REGION Network 2: Converstion all data to string
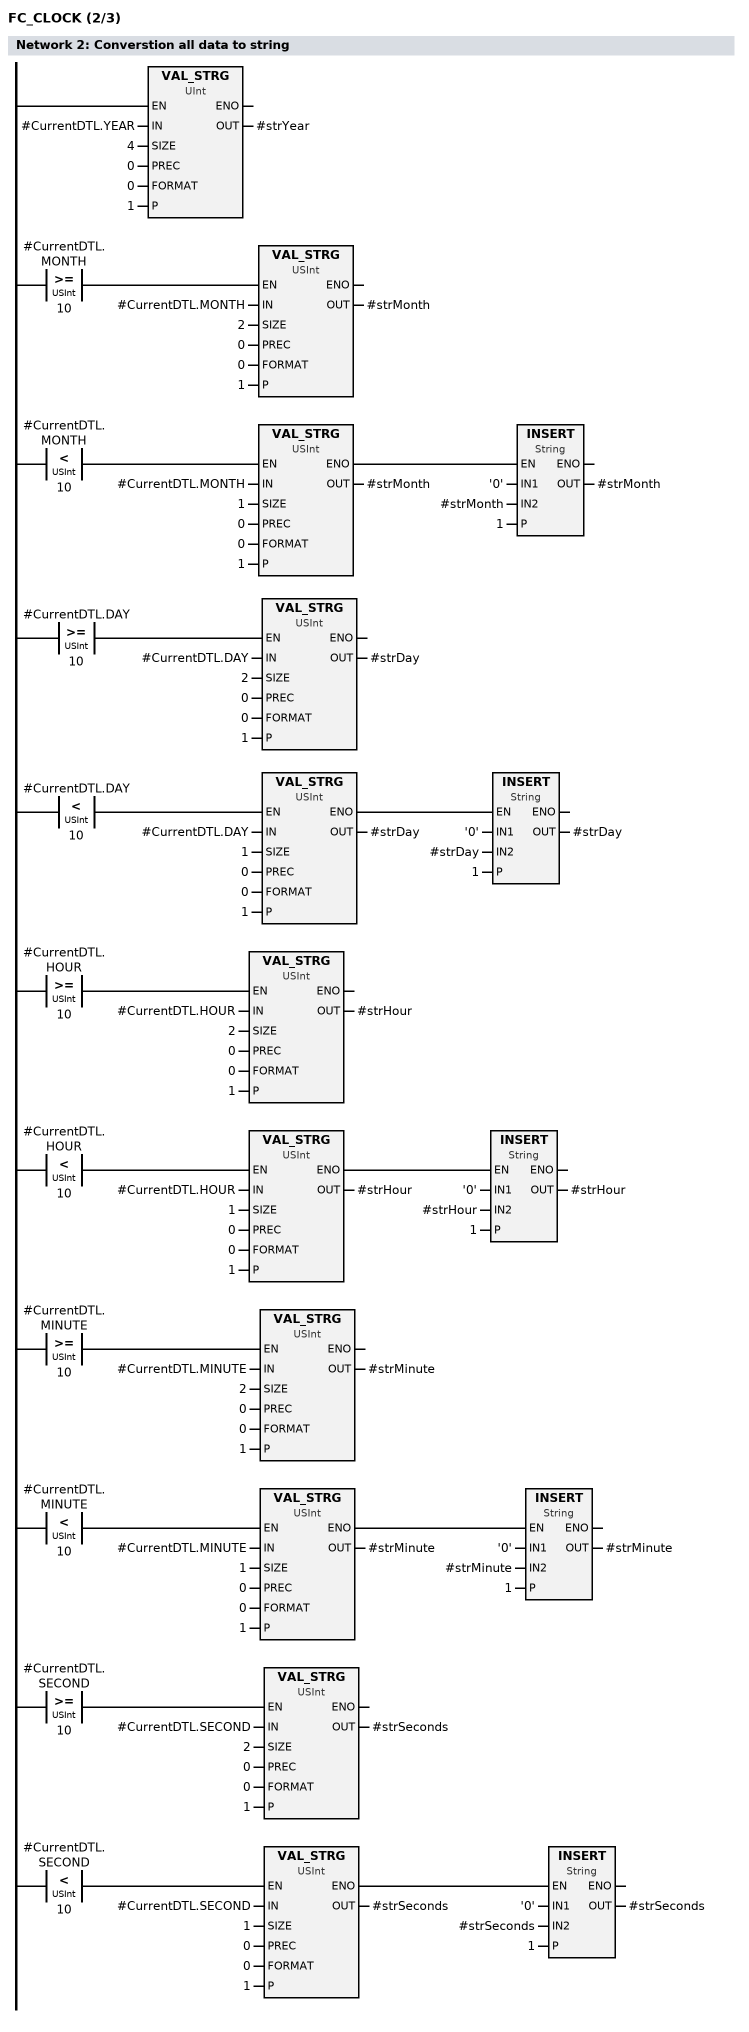
   RUNG wire#powerrail
      { S7_Templates := "[value_type := UInt, str_type := String]" } VAL_STRG(IN := #CurrentDTL.YEAR, SIZE := 4, PREC := 0, FORMAT := 0, P := 1, OUT => #strYear)
   END_RUNG
   RUNG wire#powerrail
      { S7_Templates := "SrcType := USInt" } GE_Contact(in1 := #CurrentDTL.MONTH, in2 := 10)
      { S7_Templates := "[value_type := USInt, str_type := String]" } VAL_STRG(IN := #CurrentDTL.MONTH, SIZE := 2, PREC := 0, FORMAT := 0, P := 1, OUT => #strMonth)
   END_RUNG
   RUNG wire#powerrail
      { S7_Templates := "SrcType := USInt" } LT_Contact(in1 := #CurrentDTL.MONTH, in2 := 10)
      { S7_Templates := "[value_type := USInt, str_type := String]" } VAL_STRG(IN := #CurrentDTL.MONTH, SIZE := 1, PREC := 0, FORMAT := 0, P := 1, OUT => #strMonth)
      { S7_Templates := "str_type := String" } INSERT(IN1 := '0', IN2 := #strMonth, P := 1, OUT => #strMonth)
   END_RUNG
   RUNG wire#powerrail
      { S7_Templates := "SrcType := USInt" } GE_Contact(in1 := #CurrentDTL.DAY, in2 := 10)
      { S7_Templates := "[value_type := USInt, str_type := String]" } VAL_STRG(IN := #CurrentDTL.DAY, SIZE := 2, PREC := 0, FORMAT := 0, P := 1, OUT => #strDay)
   END_RUNG
   RUNG wire#powerrail
      { S7_Templates := "SrcType := USInt" } LT_Contact(in1 := #CurrentDTL.DAY, in2 := 10)
      { S7_Templates := "[value_type := USInt, str_type := String]" } VAL_STRG(IN := #CurrentDTL.DAY, SIZE := 1, PREC := 0, FORMAT := 0, P := 1, OUT => #strDay)
      { S7_Templates := "str_type := String" } INSERT(IN1 := '0', IN2 := #strDay, P := 1, OUT => #strDay)
   END_RUNG
   RUNG wire#powerrail
      { S7_Templates := "SrcType := USInt" } GE_Contact(in1 := #CurrentDTL.HOUR, in2 := 10)
      { S7_Templates := "[value_type := USInt, str_type := String]" } VAL_STRG(IN := #CurrentDTL.HOUR, SIZE := 2, PREC := 0, FORMAT := 0, P := 1, OUT => #strHour)
   END_RUNG
   RUNG wire#powerrail
      { S7_Templates := "SrcType := USInt" } LT_Contact(in1 := #CurrentDTL.HOUR, in2 := 10)
      { S7_Templates := "[value_type := USInt, str_type := String]" } VAL_STRG(IN := #CurrentDTL.HOUR, SIZE := 1, PREC := 0, FORMAT := 0, P := 1, OUT => #strHour)
      { S7_Templates := "str_type := String" } INSERT(IN1 := '0', IN2 := #strHour, P := 1, OUT => #strHour)
   END_RUNG
   RUNG wire#powerrail
      { S7_Templates := "SrcType := USInt" } GE_Contact(in1 := #CurrentDTL.MINUTE, in2 := 10)
      { S7_Templates := "[value_type := USInt, str_type := String]" } VAL_STRG(IN := #CurrentDTL.MINUTE, SIZE := 2, PREC := 0, FORMAT := 0, P := 1, OUT => #strMinute)
   END_RUNG
   RUNG wire#powerrail
      { S7_Templates := "SrcType := USInt" } LT_Contact(in1 := #CurrentDTL.MINUTE, in2 := 10)
      { S7_Templates := "[value_type := USInt, str_type := String]" } VAL_STRG(IN := #CurrentDTL.MINUTE, SIZE := 1, PREC := 0, FORMAT := 0, P := 1, OUT => #strMinute)
      { S7_Templates := "str_type := String" } INSERT(IN1 := '0', IN2 := #strMinute, P := 1, OUT => #strMinute)
   END_RUNG
   RUNG wire#powerrail
      { S7_Templates := "SrcType := USInt" } GE_Contact(in1 := #CurrentDTL.SECOND, in2 := 10)
      { S7_Templates := "[value_type := USInt, str_type := String]" } VAL_STRG(IN := #CurrentDTL.SECOND, SIZE := 2, PREC := 0, FORMAT := 0, P := 1, OUT => #strSeconds)
   END_RUNG
   RUNG wire#powerrail
      { S7_Templates := "SrcType := USInt" } LT_Contact(in1 := #CurrentDTL.SECOND, in2 := 10)
      { S7_Templates := "[value_type := USInt, str_type := String]" } VAL_STRG(IN := #CurrentDTL.SECOND, SIZE := 1, PREC := 0, FORMAT := 0, P := 1, OUT => #strSeconds)
      { S7_Templates := "str_type := String" } INSERT(IN1 := '0', IN2 := #strSeconds, P := 1, OUT => #strSeconds)
   END_RUNG
   // the same network as SCL:
   VAL_STRG(IN := #CurrentDTL.YEAR, SIZE := 4, PREC := 0, FORMAT := 0, P := 1, OUT => #strYear);
   IF #CurrentDTL.MONTH >= 10 THEN
       VAL_STRG(IN := #CurrentDTL.MONTH, SIZE := 2, PREC := 0, FORMAT := 0, P := 1, OUT => #strMonth);
   END_IF;
   VAL_STRG(EN := #CurrentDTL.MONTH < 10,
            IN := #CurrentDTL.MONTH,
            SIZE := 1,
            PREC := 0,
            FORMAT := 0,
            P := 1,
            OUT => #strMonth,
            ENO => #_w1);
   IF #_w1 THEN INSERT(IN1 := '0', IN2 := #strMonth, P := 1, OUT => #strMonth); END_IF;
   IF #CurrentDTL.DAY >= 10 THEN
       VAL_STRG(IN := #CurrentDTL.DAY, SIZE := 2, PREC := 0, FORMAT := 0, P := 1, OUT => #strDay);
   END_IF;
   VAL_STRG(EN := #CurrentDTL.DAY < 10,
            IN := #CurrentDTL.DAY,
            SIZE := 1,
            PREC := 0,
            FORMAT := 0,
            P := 1,
            OUT => #strDay,
            ENO => #_w2);
   IF #_w2 THEN INSERT(IN1 := '0', IN2 := #strDay, P := 1, OUT => #strDay); END_IF;
   IF #CurrentDTL.HOUR >= 10 THEN
       VAL_STRG(IN := #CurrentDTL.HOUR, SIZE := 2, PREC := 0, FORMAT := 0, P := 1, OUT => #strHour);
   END_IF;
   VAL_STRG(EN := #CurrentDTL.HOUR < 10,
            IN := #CurrentDTL.HOUR,
            SIZE := 1,
            PREC := 0,
            FORMAT := 0,
            P := 1,
            OUT => #strHour,
            ENO => #_w3);
   IF #_w3 THEN INSERT(IN1 := '0', IN2 := #strHour, P := 1, OUT => #strHour); END_IF;
   IF #CurrentDTL.MINUTE >= 10 THEN
       VAL_STRG(IN := #CurrentDTL.MINUTE, SIZE := 2, PREC := 0, FORMAT := 0, P := 1, OUT => #strMinute);
   END_IF;
   VAL_STRG(EN := #CurrentDTL.MINUTE < 10,
            IN := #CurrentDTL.MINUTE,
            SIZE := 1,
            PREC := 0,
            FORMAT := 0,
            P := 1,
            OUT => #strMinute,
            ENO => #_w4);
   IF #_w4 THEN INSERT(IN1 := '0', IN2 := #strMinute, P := 1, OUT => #strMinute); END_IF;
   IF #CurrentDTL.SECOND >= 10 THEN
       VAL_STRG(IN := #CurrentDTL.SECOND, SIZE := 2, PREC := 0, FORMAT := 0, P := 1, OUT => #strSeconds);
   END_IF;
   VAL_STRG(EN := #CurrentDTL.SECOND < 10,
            IN := #CurrentDTL.SECOND,
            SIZE := 1,
            PREC := 0,
            FORMAT := 0,
            P := 1,
            OUT => #strSeconds,
            ENO => #_w5);
   IF #_w5 THEN INSERT(IN1 := '0', IN2 := #strSeconds, P := 1, OUT => #strSeconds); END_IF;
END_REGION

REGION Network 3: Current Time String
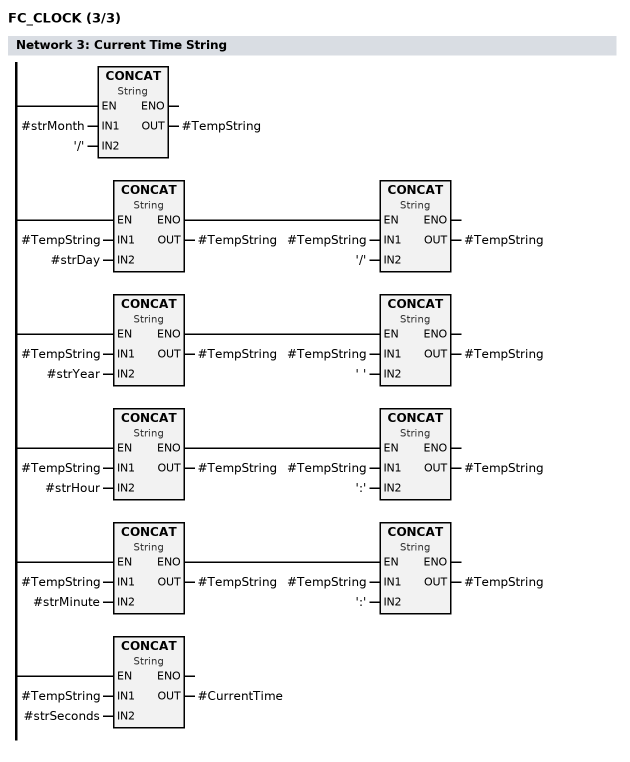
   RUNG wire#powerrail
      { S7_Templates := "[card := 2, str_type := String]" } CONCAT(IN1 := #strMonth, IN2 := '/', OUT => #TempString)
   END_RUNG
   RUNG wire#powerrail
      { S7_Templates := "[card := 2, str_type := String]" } CONCAT(IN1 := #TempString, IN2 := #strDay, OUT => #TempString)
      { S7_Templates := "[card := 2, str_type := String]" } CONCAT(IN1 := #TempString, IN2 := '/', OUT => #TempString)
   END_RUNG
   RUNG wire#powerrail
      { S7_Templates := "[card := 2, str_type := String]" } CONCAT(IN1 := #TempString, IN2 := #strYear, OUT => #TempString)
      { S7_Templates := "[card := 2, str_type := String]" } CONCAT(IN1 := #TempString, IN2 := ' ', OUT => #TempString)
   END_RUNG
   RUNG wire#powerrail
      { S7_Templates := "[card := 2, str_type := String]" } CONCAT(IN1 := #TempString, IN2 := #strHour, OUT => #TempString)
      { S7_Templates := "[card := 2, str_type := String]" } CONCAT(IN1 := #TempString, IN2 := ':', OUT => #TempString)
   END_RUNG
   RUNG wire#powerrail
      { S7_Templates := "[card := 2, str_type := String]" } CONCAT(IN1 := #TempString, IN2 := #strMinute, OUT => #TempString)
      { S7_Templates := "[card := 2, str_type := String]" } CONCAT(IN1 := #TempString, IN2 := ':', OUT => #TempString)
   END_RUNG
   RUNG wire#powerrail
      { S7_Templates := "[card := 2, str_type := String]" } CONCAT(IN1 := #TempString, IN2 := #strSeconds, OUT => #CurrentTime)
   END_RUNG
   // the same network as SCL:
   CONCAT(IN1 := #strMonth, IN2 := '/', OUT => #TempString);
   CONCAT(IN1 := #TempString, IN2 := #strDay, OUT => #TempString, ENO => #_w1);
   IF #_w1 THEN CONCAT(IN1 := #TempString, IN2 := '/', OUT => #TempString); END_IF;
   CONCAT(IN1 := #TempString, IN2 := #strYear, OUT => #TempString, ENO => #_w2);
   IF #_w2 THEN CONCAT(IN1 := #TempString, IN2 := ' ', OUT => #TempString); END_IF;
   CONCAT(IN1 := #TempString, IN2 := #strHour, OUT => #TempString, ENO => #_w3);
   IF #_w3 THEN CONCAT(IN1 := #TempString, IN2 := ':', OUT => #TempString); END_IF;
   CONCAT(IN1 := #TempString, IN2 := #strMinute, OUT => #TempString, ENO => #_w4);
   IF #_w4 THEN CONCAT(IN1 := #TempString, IN2 := ':', OUT => #TempString); END_IF;
   CONCAT(IN1 := #TempString, IN2 := #strSeconds, OUT => #CurrentTime);
END_REGION
END_FUNCTION

FUNCTION_BLOCK "FB_HeartBeat"   // FB25, SCL
{ S7_Optimized_Access := 'TRUE' }
VERSION : 0.1
// stored: AutoNumber true, IsIECCheckEnabled false, IsRetainMemResEnabled false, MemoryReserve 100, SetENOAutomatically false, UDAEnableTagReadback false
   VAR_INPUT
      PC_HeartBeat : Word;
   END_VAR
   VAR_OUTPUT
      PLC_HeartBeat : Word;
      PC_Disconnected : Bool;
   END_VAR
   VAR
      TimeOut : TON_TIME;
      "Timer" { S7_SetPoint := 'True'} : TON_TIME;
      PC_Heartbeat_old : Word;
      StartTimerBit : Bool := FALSE;
   END_VAR
BEGIN
   #Timer(IN := #StartTimerBit, //
          PT := t#250ms);
   IF NOT #StartTimerBit THEN
       #StartTimerBit := TRUE;
   END_IF;
   #Timer(IN := #StartTimerBit, //
          PT := t#250ms);
   IF #Timer.Q THEN
       #StartTimerBit := FALSE;
       RESET_TIMER(#Timer);
       #PLC_HeartBeat += 1;
   END_IF;
   //Time Out Timer
   #TimeOut(IN := #PC_HeartBeat = #PC_Heartbeat_old,
            PT := t#10s);
   #PC_Heartbeat_old := #PC_HeartBeat;
   #PC_Disconnected := #TimeOut.Q; // if time out set PC_Disconnected
END_FUNCTION_BLOCK

FUNCTION "OUTPUTS" : Void   // FC5, SCL
{ S7_Optimized_Access := 'TRUE' }
VERSION : 0.1
// stored: AutoNumber true, IsIECCheckEnabled false, SetENOAutomatically false, UDAEnableTagReadback false
BEGIN
   REGION MAIN PANEL
       "MAIN PANEL STACK LIGHT RED" := "Stack_Lights_DB_0".Red XOR "Force"."MAIN PANEL STACK LIGHT RED";
       "MAIN PANEL STACK LIGHT AMBER" := "Stack_Lights_DB_0".Yellow XOR "Force"."MAIN PANEL STACK LIGHT AMBER";
       "MAIN PANEL STACK LIGHT GREEN" := "Stack_Lights_DB_0".Green XOR "Force"."MAIN PANEL STACK LIGHT GREEN";
   END_REGION

   REGION REMOTE PANEL 1
       "C1101_SFTY STOPPER ROTATE" := "Sf_C1101_FB_DB".T_Run.Q XOR "Force".Remote_Panel[1]."CX101_SFTY STOPPER ROTATE";
       "C1102_SFTY STOPPER ROTATE" := "Sf_C1102_FB_DB".T_Run.Q XOR "Force".Remote_Panel[1]."CX102_SFTY STOPPER ROTATE";
       "C1103_SFTY STOPPER ROTATE" := "Sf_C1103_FB_DB".T_Run.Q XOR "Force".Remote_Panel[1]."CX103_SFTY STOPPER ROTATE";
       "C1104_SFTY STOPPER ROTATE" := "Sf_C1104_FB_DB".T_Run.Q XOR "Force".Remote_Panel[1]."CX104_SFTY STOPPER ROTATE";
       "C1105_SFTY STOPPER ROTATE" := "Sf_C1105_FB_DB".T_Run.Q XOR "Force".Remote_Panel[1]."CX105_SFTY STOPPER ROTATE";
       "C1106_SFTY STOPPER ROTATE" := "Sf_C1106_FB_DB".T_Run.Q XOR "Force".Remote_Panel[1]."CX106_SFTY STOPPER ROTATE";
       "C1107_SFTY STOPPER ROTATE" := "Sf_C1107_FB_DB".T_Run.Q XOR "Force".Remote_Panel[1]."CX107_SFTY STOPPER ROTATE";
       "C1108_SFTY STOPPER ROTATE" := "Sf_C1108_FB_DB".T_Run.Q XOR "Force".Remote_Panel[1]."CX108_SFTY STOPPER ROTATE";
       "C1201_SFTY STOPPER ROTATE" := "Sf_C1201_FB_DB".T_Run.Q XOR "Force".Remote_Panel[1]."CX201_SFTY STOPPER ROTATE";
       "C1202_SFTY STOPPER ROTATE" := "Sf_C1202_FB_DB".T_Run.Q XOR "Force".Remote_Panel[1]."CX202_SFTY STOPPER ROTATE";
       "C1203_SFTY STOPPER ROTATE" := "Sf_C1203_FB_DB".T_Run.Q XOR "Force".Remote_Panel[1]."CX203_SFTY STOPPER ROTATE";
       "C1204_SFTY STOPPER ROTATE" := "Sf_C1204_FB_DB".T_Run.Q XOR "Force".Remote_Panel[1]."CX204_SFTY STOPPER ROTATE";
       "C1205_SFTY STOPPER ROTATE" := "Sf_C1205_FB_DB".T_Run.Q XOR "Force".Remote_Panel[1]."CX205_SFTY STOPPER ROTATE";
       "C1206_SFTY STOPPER ROTATE" := "Sf_C1206_FB_DB".T_Run.Q XOR "Force".Remote_Panel[1]."CX206_SFTY STOPPER ROTATE";
       "C1207_SFTY STOPPER ROTATE" := "Sf_C1207_FB_DB".T_Run.Q XOR "Force".Remote_Panel[1]."CX207_SFTY STOPPER ROTATE";
       "C1208_SFTY STOPPER ROTATE" := "Sf_C1208_FB_DB".T_Run.Q XOR "Force".Remote_Panel[1]."CX208_SFTY STOPPER ROTATE";
       "VTD1 DOCKING PINS 1 EXTEND" := "Control_DB".VTD_Sys[1].Outputs.LP1_Extend XOR "Force".Remote_Panel[1]."VTDx DOCKING PINS 1 EXTEND";
       "VTD1 DOCKING PINS 1 RETRACT" := "Control_DB".VTD_Sys[1].Outputs.LP1_Retract XOR "Force".Remote_Panel[1]."VTDx DOCKING PINS 1 RETRACT";
       "VTD1 DOCKING PINS 2 EXTEND" := "Control_DB".VTD_Sys[1].Outputs.LP2_Extend XOR "Force".Remote_Panel[1]."VTDx DOCKING PINS 2 EXTEND";
       "VTD1 DOCKING PINS 2 RETRACT" := "Control_DB".VTD_Sys[1].Outputs.LP2_Retract XOR "Force".Remote_Panel[1]."VTDx DOCKING PINS 2 RETRACT";
       "SCA 1002 STACK LIGHTS AMBER" := "Stack_Lights_DB_1".Yellow XOR "Force".Remote_Panel[1]."SCA X00Y STACK LIGHTS AMBER";
       "SCA 1002 STACK LIGHTS GREEN" := "Stack_Lights_DB_1".Green XOR "Force".Remote_Panel[1]."SCA X00Y STACK LIGHTS GREEN";
       "SCA 1002 STACK LIGHTS RED" := "Stack_Lights_DB_1".Red XOR "Force".Remote_Panel[1]."SCA X00Y STACK LIGHTS RED";
       "EMERGENCY STOP RESET STATUS - ON(1)" := "Force".Remote_Panel[1]."EMERGENCY STOP RESET STATUS - ON(X)" XOR (NOT "Remote_Panel_DB_1".Safety_OK AND "Clock_2Hz");

       "VTD1_ControlWord".%X7 := "Control_DB".VTD_Sys[1].Instruction.Reset;
       "VTD1_AccFactor" := "Control_DB".VTD_Sys[1].Motor.Acc_Factor;

       //ABSOLUTE ENMCODER
       "AE_Control_Word_1(1)" := "Control_DB".VTD_Sys[1].Outputs.AE_Control_Word_1;
       "AE_Control_Word_2(1)" := "Control_DB".VTD_Sys[1].Outputs.AE_Control_Word_2;
   END_REGION

   REGION REMOTE PANEL 2
       "C2101_SFTY STOPPER ROTATE" := "Sf_C2101_FB_DB".T_Run.Q XOR "Force".Remote_Panel[2]."CX101_SFTY STOPPER ROTATE";
       "C2102_SFTY STOPPER ROTATE" := "Sf_C2102_FB_DB".T_Run.Q XOR "Force".Remote_Panel[2]."CX102_SFTY STOPPER ROTATE";
       "C2103_SFTY STOPPER ROTATE" := "Sf_C2103_FB_DB".T_Run.Q XOR "Force".Remote_Panel[2]."CX103_SFTY STOPPER ROTATE";
       "C2104_SFTY STOPPER ROTATE" := "Sf_C2104_FB_DB".T_Run.Q XOR "Force".Remote_Panel[2]."CX104_SFTY STOPPER ROTATE";
       "C2105_SFTY STOPPER ROTATE" := "Sf_C2105_FB_DB".T_Run.Q XOR "Force".Remote_Panel[2]."CX105_SFTY STOPPER ROTATE";
       "C2106_SFTY STOPPER ROTATE" := "Sf_C2106_FB_DB".T_Run.Q XOR "Force".Remote_Panel[2]."CX106_SFTY STOPPER ROTATE";
       "C2107_SFTY STOPPER ROTATE" := "Sf_C2107_FB_DB".T_Run.Q XOR "Force".Remote_Panel[2]."CX107_SFTY STOPPER ROTATE";
       "C2108_SFTY STOPPER ROTATE" := "Sf_C2108_FB_DB".T_Run.Q XOR "Force".Remote_Panel[2]."CX108_SFTY STOPPER ROTATE";
       "C2201_SFTY STOPPER ROTATE" := "Sf_C2201_FB_DB".T_Run.Q XOR "Force".Remote_Panel[2]."CX201_SFTY STOPPER ROTATE";
       "C2202_SFTY STOPPER ROTATE" := "Sf_C2202_FB_DB".T_Run.Q XOR "Force".Remote_Panel[2]."CX202_SFTY STOPPER ROTATE";
       "C2203_SFTY STOPPER ROTATE" := "Sf_C2203_FB_DB".T_Run.Q XOR "Force".Remote_Panel[2]."CX203_SFTY STOPPER ROTATE";
       "C2204_SFTY STOPPER ROTATE" := "Sf_C2204_FB_DB".T_Run.Q XOR "Force".Remote_Panel[2]."CX204_SFTY STOPPER ROTATE";
       "C2205_SFTY STOPPER ROTATE" := "Sf_C2205_FB_DB".T_Run.Q XOR "Force".Remote_Panel[2]."CX205_SFTY STOPPER ROTATE";
       "C2206_SFTY STOPPER ROTATE" := "Sf_C2206_FB_DB".T_Run.Q XOR "Force".Remote_Panel[2]."CX206_SFTY STOPPER ROTATE";
       "C2207_SFTY STOPPER ROTATE" := "Sf_C2207_FB_DB".T_Run.Q XOR "Force".Remote_Panel[2]."CX207_SFTY STOPPER ROTATE";
       "C2208_SFTY STOPPER ROTATE" := "Sf_C2208_FB_DB".T_Run.Q XOR "Force".Remote_Panel[2]."CX208_SFTY STOPPER ROTATE";
       "VTD2 DOCKING PINS 1 EXTEND" := "Control_DB".VTD_Sys[2].Outputs.LP1_Extend XOR "Force".Remote_Panel[2]."VTDx DOCKING PINS 1 EXTEND";
       "VTD2 DOCKING PINS 1 RETRACT" := "Control_DB".VTD_Sys[2].Outputs.LP1_Retract XOR "Force".Remote_Panel[2]."VTDx DOCKING PINS 1 RETRACT";
       "VTD2 DOCKING PINS 2 EXTEND" := "Control_DB".VTD_Sys[2].Outputs.LP2_Extend XOR "Force".Remote_Panel[2]."VTDx DOCKING PINS 2 EXTEND";
       "VTD2 DOCKING PINS 2 RETRACT" := "Control_DB".VTD_Sys[2].Outputs.LP2_Retract XOR "Force".Remote_Panel[2]."VTDx DOCKING PINS 2 RETRACT";
       "SCA 2002 STACK LIGHTS AMBER" := "Stack_Lights_DB_2".Yellow XOR "Force".Remote_Panel[2]."SCA X00Y STACK LIGHTS AMBER";
       "SCA 2002 STACK LIGHTS RED" := "Stack_Lights_DB_2".Red XOR "Force".Remote_Panel[2]."SCA X00Y STACK LIGHTS RED";
       "SCA 2002 STACK LIGHTS GREEN" := "Stack_Lights_DB_2".Green XOR "Force".Remote_Panel[2]."SCA X00Y STACK LIGHTS GREEN";
       "EMERGENCY STOP RESET STATUS - ON(2)" := "Force".Remote_Panel[2]."EMERGENCY STOP RESET STATUS - ON(X)" XOR (NOT "Remote_Panel_DB_2".Safety_OK AND "Clock_2Hz");

       "VTD2_ControlWord".%X7 := "Control_DB".VTD_Sys[2].Instruction.Reset;
       "VTD2_AccFactor" := "Control_DB".VTD_Sys[2].Motor.Acc_Factor;

       //ABSOLUTE ENMCODER
       "AE_Control_Word_1(2)" := "Control_DB".VTD_Sys[2].Outputs.AE_Control_Word_1;
       "AE_Control_Word_2(2)" := "Control_DB".VTD_Sys[2].Outputs.AE_Control_Word_2;
   END_REGION

   REGION REMOTE PANEL 3
       "C3101_SFTY STOPPER ROTATE" := "Sf_C3101_FB_DB".T_Run.Q XOR "Force".Remote_Panel[3]."CX101_SFTY STOPPER ROTATE";
       "C3102_SFTY STOPPER ROTATE" := "Sf_C3102_FB_DB".T_Run.Q XOR "Force".Remote_Panel[3]."CX102_SFTY STOPPER ROTATE";
       "C3103_SFTY STOPPER ROTATE" := "Sf_C3103_FB_DB".T_Run.Q XOR "Force".Remote_Panel[3]."CX103_SFTY STOPPER ROTATE";
       "C3104_SFTY STOPPER ROTATE" := "Sf_C3104_FB_DB".T_Run.Q XOR "Force".Remote_Panel[3]."CX104_SFTY STOPPER ROTATE";
       "C3105_SFTY STOPPER ROTATE" := "Sf_C3105_FB_DB".T_Run.Q XOR "Force".Remote_Panel[3]."CX105_SFTY STOPPER ROTATE";
       "C3106_SFTY STOPPER ROTATE" := "Sf_C3106_FB_DB".T_Run.Q XOR "Force".Remote_Panel[3]."CX106_SFTY STOPPER ROTATE";
       "C3107_SFTY STOPPER ROTATE" := "Sf_C3107_FB_DB".T_Run.Q XOR "Force".Remote_Panel[3]."CX107_SFTY STOPPER ROTATE";
       "C3108_SFTY STOPPER ROTATE" := "Sf_C3108_FB_DB".T_Run.Q XOR "Force".Remote_Panel[3]."CX208_SFTY STOPPER ROTATE";
       "C3201_SFTY STOPPER ROTATE" := "Sf_C3201_FB_DB".T_Run.Q XOR "Force".Remote_Panel[3]."CX201_SFTY STOPPER ROTATE";
       "C3202_SFTY STOPPER ROTATE" := "Sf_C3202_FB_DB".T_Run.Q XOR "Force".Remote_Panel[3]."CX202_SFTY STOPPER ROTATE";
       "C3203_SFTY STOPPER ROTATE" := "Sf_C3203_FB_DB".T_Run.Q XOR "Force".Remote_Panel[3]."CX203_SFTY STOPPER ROTATE";
       "C3204_SFTY STOPPER ROTATE" := "Sf_C3204_FB_DB".T_Run.Q XOR "Force".Remote_Panel[3]."CX204_SFTY STOPPER ROTATE";
       "C3205_SFTY STOPPER ROTATE" := "Sf_C3205_FB_DB".T_Run.Q XOR "Force".Remote_Panel[3]."CX205_SFTY STOPPER ROTATE";
       "C3206_SFTY STOPPER ROTATE" := "Sf_C3206_FB_DB".T_Run.Q XOR "Force".Remote_Panel[3]."CX206_SFTY STOPPER ROTATE";
       "C3207_SFTY STOPPER ROTATE" := "Sf_C3207_FB_DB".T_Run.Q XOR "Force".Remote_Panel[3]."CX207_SFTY STOPPER ROTATE";
       "C3208_SFTY STOPPER ROTATE" := "Sf_C3208_FB_DB".T_Run.Q XOR "Force".Remote_Panel[3]."CX208_SFTY STOPPER ROTATE";
       "VTD3 DOCKING PINS 1 EXTEND" := "Control_DB".VTD_Sys[3].Outputs.LP1_Extend XOR "Force".Remote_Panel[3]."VTDx DOCKING PINS 1 EXTEND";
       "VTD3 DOCKING PINS 1 RETRACT" := "Control_DB".VTD_Sys[3].Outputs.LP1_Retract XOR "Force".Remote_Panel[3]."VTDx DOCKING PINS 1 RETRACT";
       "VTD3 DOCKING PINS 2 EXTEND" := "Control_DB".VTD_Sys[3].Outputs.LP2_Extend XOR "Force".Remote_Panel[3]."VTDx DOCKING PINS 2 EXTEND";
       "VTD3 DOCKING PINS 2 RETRACT" := "Control_DB".VTD_Sys[3].Outputs.LP2_Retract XOR "Force".Remote_Panel[3]."VTDx DOCKING PINS 2 RETRACT";
       "SCA 3002 STACK LIGHTS RED" := "Stack_Lights_DB_3".Red XOR "Force".Remote_Panel[3]."SCA X00Y STACK LIGHTS RED";
       "SCA 3002 STACK LIGHTS ORANGE" := "Stack_Lights_DB_3".Yellow XOR "Force".Remote_Panel[3]."SCA X00Y STACK LIGHTS AMBER";
       "SCA 3002 STACK LIGHTS GREEN" := "Stack_Lights_DB_3".Green XOR "Force".Remote_Panel[3]."SCA X00Y STACK LIGHTS GREEN";
       "EMERGENCY STOP RESET STATUS - ON(3)" := "Force".Remote_Panel[3]."EMERGENCY STOP RESET STATUS - ON(X)" XOR (NOT "Remote_Panel_DB_3".Safety_OK AND "Clock_2Hz");

       "VTD3_ControlWord".%X7 := "Control_DB".VTD_Sys[3].Instruction.Reset;
       "VTD3_AccFactor" := "Control_DB".VTD_Sys[3].Motor.Acc_Factor;

       //ABSOLUTE ENMCODER
       "AE_Control_Word_1(3)" := "Control_DB".VTD_Sys[3].Outputs.AE_Control_Word_1;
       "AE_Control_Word_2(3)" := "Control_DB".VTD_Sys[3].Outputs.AE_Control_Word_2;
   END_REGION

   REGION REMOTE PANEL 4
       "C4101_SFTY STOPPER ROTATE" := "Sf_C4101_FB_DB".T_Run.Q XOR "Force".Remote_Panel[4]."CX101_SFTY STOPPER ROTATE";
       "C4102_SFTY STOPPER ROTATE" := "Sf_C4102_FB_DB".T_Run.Q XOR "Force".Remote_Panel[4]."CX102_SFTY STOPPER ROTATE";
       "C4103_SFTY STOPPER ROTATE" := "Sf_C4103_FB_DB".T_Run.Q XOR "Force".Remote_Panel[4]."CX103_SFTY STOPPER ROTATE";
       "C4104_SFTY STOPPER ROTATE" := "Sf_C4104_FB_DB".T_Run.Q XOR "Force".Remote_Panel[4]."CX104_SFTY STOPPER ROTATE";
       "C4105_SFTY STOPPER ROTATE" := "Sf_C4105_FB_DB".T_Run.Q XOR "Force".Remote_Panel[4]."CX105_SFTY STOPPER ROTATE";
       "C4106_SFTY STOPPER ROTATE" := "Sf_C4106_FB_DB".T_Run.Q XOR "Force".Remote_Panel[4]."CX106_SFTY STOPPER ROTATE";
       "C4107_SFTY STOPPER ROTATE" := "Sf_C4107_FB_DB".T_Run.Q XOR "Force".Remote_Panel[4]."CX107_SFTY STOPPER ROTATE";
       "C4108_SFTY STOPPER ROTATE" := "Sf_C4108_FB_DB".T_Run.Q XOR "Force".Remote_Panel[4]."CX108_SFTY STOPPER ROTATE";
       "VTD4 DOCKING PINS 1 EXTEND" := "Control_DB".VTD_Sys[4].Outputs.LP1_Extend XOR "Force".Remote_Panel[4]."VTDx DOCKING PINS 1 EXTEND";
       "VTD4 DOCKING PINS 1 RETRACT" := "Control_DB".VTD_Sys[4].Outputs.LP1_Retract XOR "Force".Remote_Panel[4]."VTDx DOCKING PINS 1 RETRACT";
       "VTD4 DOCKING PINS 2 EXTEND" := "Control_DB".VTD_Sys[4].Outputs.LP2_Extend XOR "Force".Remote_Panel[4]."VTDx DOCKING PINS 2 EXTEND";
       "VTD4 DOCKING PINS 2 RETRACT" := "Control_DB".VTD_Sys[4].Outputs.LP2_Retract XOR "Force".Remote_Panel[4]."VTDx DOCKING PINS 2 RETRACT";
       "SCA 4001 STACK LIGHTS RED" := "Stack_Lights_DB_4".Red XOR "Force".Remote_Panel[4]."SCA X00Y STACK LIGHTS RED";
       "SCA 4001 STACK LIGHTS YELLOW" := "Stack_Lights_DB_4".Yellow XOR "Force".Remote_Panel[4]."SCA X00Y STACK LIGHTS AMBER";
       "SCA 4001 STACK LIGHTS GREEN" := "Stack_Lights_DB_4".Green XOR "Force".Remote_Panel[4]."SCA X00Y STACK LIGHTS GREEN";
       "EMERGENCY STOP RESET STATUS - ON(4)" := "Force".Remote_Panel[4]."EMERGENCY STOP RESET STATUS - ON(X)" XOR (NOT "Remote_Panel_DB_4".Safety_OK AND "Clock_2Hz");

       "VTD4_ControlWord".%X7 := "Control_DB".VTD_Sys[4].Instruction.Reset;
       "VTD4_AccFactor" := "Control_DB".VTD_Sys[4].Motor.Acc_Factor;

       //ABSOLUTE ENMCODER
       "AE_Control_Word_1(4)" := "Control_DB".VTD_Sys[4].Outputs.AE_Control_Word_1;
       "AE_Control_Word_2(4)" := "Control_DB".VTD_Sys[4].Outputs.AE_Control_Word_2;
   END_REGION

   REGION REMOTE PANEL 5
       "C5101_SFTY STOPPER ROTATE" := "Sf_C5101_FB_DB".T_Run.Q XOR "Force".Remote_Panel[5]."CX101_SFTY STOPPER ROTATE";
       "C5102_SFTY STOPPER ROTATE" := "Sf_C5102_FB_DB".T_Run.Q XOR "Force".Remote_Panel[5]."CX102_SFTY STOPPER ROTATE";
       "C5103_SFTY STOPPER ROTATE" := "Sf_C5103_FB_DB".T_Run.Q XOR "Force".Remote_Panel[5]."CX103_SFTY STOPPER ROTATE";
       "C5104_SFTY STOPPER ROTATE" := "Sf_C5104_FB_DB".T_Run.Q XOR "Force".Remote_Panel[5]."CX104_SFTY STOPPER ROTATE";
       "C5105_SFTY STOPPER ROTATE" := "Sf_C5105_FB_DB".T_Run.Q XOR "Force".Remote_Panel[5]."CX105_SFTY STOPPER ROTATE";
       "C5106_SFTY STOPPER ROTATE" := "Sf_C5106_FB_DB".T_Run.Q XOR "Force".Remote_Panel[5]."CX106_SFTY STOPPER ROTATE";
       "C5107_SFTY STOPPER ROTATE" := "Sf_C5107_FB_DB".T_Run.Q XOR "Force".Remote_Panel[5]."CX107_SFTY STOPPER ROTATE";
       "C5108_SFTY STOPPER ROTATE" := "Sf_C5108_FB_DB".T_Run.Q XOR "Force".Remote_Panel[5]."CX108_SFTY STOPPER ROTATE";
       "VTD5 DOCKING PINS 1 EXTEND" := "Control_DB".VTD_Sys[5].Outputs.LP1_Extend XOR "Force".Remote_Panel[5]."VTDx DOCKING PINS 1 EXTEND";
       "VTD5 DOCKING PINS 1 RETRACT" := "Control_DB".VTD_Sys[5].Outputs.LP1_Retract XOR "Force".Remote_Panel[5]."VTDx DOCKING PINS 1 RETRACT";
       "VTD5 DOCKING PINS 2 EXTEND" := "Control_DB".VTD_Sys[5].Outputs.LP2_Extend XOR "Force".Remote_Panel[5]."VTDx DOCKING PINS 2 EXTEND";
       "VTD5 DOCKING PINS 2 RETRACT" := "Control_DB".VTD_Sys[5].Outputs.LP2_Retract XOR "Force".Remote_Panel[5]."VTDx DOCKING PINS 2 RETRACT";
       "SCA 5001 STACK LIGHTS GREEN" := "Stack_Lights_DB_5".Green XOR "Force".Remote_Panel[5]."SCA X00Y STACK LIGHTS GREEN";
       "SCA 5001 STACK LIGHTS YELLOW" := "Stack_Lights_DB_5".Yellow XOR "Force".Remote_Panel[5]."SCA X00Y STACK LIGHTS AMBER";
       "SCA 5001 STACK LIGHTS RED" := "Stack_Lights_DB_5".Red XOR "Force".Remote_Panel[5]."SCA X00Y STACK LIGHTS RED";
       "EMERGENCY STOP RESET STATUS - ON(5)" := "Force".Remote_Panel[5]."EMERGENCY STOP RESET STATUS - ON(X)" XOR (NOT "Remote_Panel_DB_5".Safety_OK AND "Clock_2Hz");

       "VTD5_ControlWord".%X7 := "Control_DB".VTD_Sys[5].Instruction.Reset;
       "VTD5_AccFactor" := "Control_DB".VTD_Sys[5].Motor.Acc_Factor;

       //ABSOLUTE ENMCODER
       "AE_Control_Word_1(5)" := "Control_DB".VTD_Sys[5].Outputs.AE_Control_Word_1;
       "AE_Control_Word_2(5)" := "Control_DB".VTD_Sys[5].Outputs.AE_Control_Word_2;
   END_REGION

   REGION CHARGER PANELS   
       IF "FirstScan" THEN
           "Charger 1 contactor(1)" := TRUE;
           "Charger 2 contactor(1)" := TRUE;
           "Charger 3 contactor(1)" := TRUE;

           "Charger 1 contactor(2)" := TRUE;
           "Charger 2 contactor(2)" := TRUE;
           "Charger 3 contactor(2)" := TRUE;

           "Charger 1 contactor(3)" := TRUE;
           "Charger 2 contactor(3)" := TRUE;
           "Charger 3 contactor(3)" := TRUE;

           "Charger 1 contactor(4)" := TRUE;
           "Charger 2 contactor(4)" := TRUE;
           "Charger 3 contactor(4)" := TRUE;

           "Charger 1 contactor(5)" := TRUE;
           "Charger 2 contactor(5)" := TRUE;
           "Charger 3 contactor(5)" := TRUE;

           "Charger 1 contactor(6)" := TRUE;
           "Charger 2 contactor(6)" := TRUE;
           "Charger 3 contactor(6)" := TRUE;

           "Charger 1 contactor(7)" := TRUE;
           "Charger 2 contactor(7)" := TRUE;
           "Charger 3 contactor(7)" := TRUE;

           "Charger 1 contactor(8)" := TRUE;
           "Charger 2 contactor(8)" := TRUE;
           "Charger 3 contactor(8)" := TRUE;

           //CHARGE DATA HMI 1
       ELSIF "Charge_Shuttle_Commands" THEN
           CASE "Shuttle_Level_Selected" OF
               1:
                   "Charger 1" := "Charger 1 contactor(1)";
                   "Charger 2" := "Charger 2 contactor(1)";
                   "Charger 3" := "Charger 3 contactor(1)";
               2:
                   "Charger 1" := "Charger 1 contactor(2)";
                   "Charger 2" := "Charger 2 contactor(2)";
                   "Charger 3" := "Charger 3 contactor(2)";
               3:
                   "Charger 1" := "Charger 1 contactor(3)";
                   "Charger 2" := "Charger 2 contactor(3)";
                   "Charger 3" := "Charger 3 contactor(3)";
               4:
                   "Charger 1" := "Charger 1 contactor(4)";
                   "Charger 2" := "Charger 2 contactor(4)";
                   "Charger 3" := "Charger 3 contactor(4)";
               5:
                   "Charger 1" := "Charger 1 contactor(5)";
                   "Charger 2" := "Charger 2 contactor(5)";
                   "Charger 3" := "Charger 3 contactor(5)";
               6:
                   "Charger 1" := "Charger 1 contactor(6)";
                   "Charger 2" := "Charger 2 contactor(6)";
                   "Charger 3" := "Charger 3 contactor(6)";
               7:
                   "Charger 1" := "Charger 1 contactor(7)";
                   "Charger 2" := "Charger 2 contactor(7)";
                   "Charger 3" := "Charger 3 contactor(7)";
               8:
                   "Charger 1" := "Charger 1 contactor(8)";
                   "Charger 2" := "Charger 2 contactor(8)";
                   "Charger 3" := "Charger 3 contactor(8)";
           END_CASE;

         "T_Shuttle_Charge_Buttons".TON(IN:=TRUE,
                                        PT:=T#100ms);

         IF "T_Shuttle_Charge_Buttons".Q THEN
             "T_Shuttle_Charge_Buttons".TON(IN := FALSE,
                                            PT := T#0S);
             "Charge_Shuttle_Commands" := FALSE;
         END_IF;

       ELSE
           //WRITE DATA
           CASE "Shuttle_Level_Selected" OF
               1:
                   "Charger 1 contactor(1)" := "Charger 1";
                   "Charger 2 contactor(1)" := "Charger 2";
                   "Charger 3 contactor(1)" := "Charger 3";
               2:
                   "Charger 1 contactor(2)" := "Charger 1";
                   "Charger 2 contactor(2)" := "Charger 2";
                   "Charger 3 contactor(2)" := "Charger 3";
               3:
                   "Charger 1 contactor(3)" := "Charger 1";
                   "Charger 2 contactor(3)" := "Charger 2";
                   "Charger 3 contactor(3)" := "Charger 3";
               4:
                   "Charger 1 contactor(4)" := "Charger 1";
                   "Charger 2 contactor(4)" := "Charger 2";
                   "Charger 3 contactor(4)" := "Charger 3";
               5:
                   "Charger 1 contactor(5)" := "Charger 1";
                   "Charger 2 contactor(5)" := "Charger 2";
                   "Charger 3 contactor(5)" := "Charger 3";
               6:
                   "Charger 1 contactor(6)" := "Charger 1";
                   "Charger 2 contactor(6)" := "Charger 2";
                   "Charger 3 contactor(6)" := "Charger 3";
               7:
                   "Charger 1 contactor(7)" := "Charger 1";
                   "Charger 2 contactor(7)" := "Charger 2";
                   "Charger 3 contactor(7)" := "Charger 3";
               8:
                   "Charger 1 contactor(8)" := "Charger 1";
                   "Charger 2 contactor(8)" := "Charger 2";
                   "Charger 3 contactor(8)" := "Charger 3";
           END_CASE;
       END_IF;
   END_REGION;
END_FUNCTION

ORGANIZATION_BLOCK "PullOrPlugOfModules"   // OB83, LAD, PullOrPlugOfModules
{ S7_Optimized_Access := 'TRUE' }
VERSION : 0.1
// stored: IsIECCheckEnabled false, SetENOAutomatically false
   VAR_INPUT
      LADDR : HW_IO;   // Hardware identifier
      Event_Class : Byte;   // 16#38/39: module inserted, removed
      Fault_ID : Byte;   // Fault identifier
   END_VAR
BEGIN
END_ORGANIZATION_BLOCK

ORGANIZATION_BLOCK "RackOrStationFailure"   // OB86, LAD, RackOrStationFailure
{ S7_Optimized_Access := 'TRUE' }
VERSION : 0.1
// stored: IsIECCheckEnabled false, SetENOAutomatically false
   VAR_INPUT
      LADDR : HW_DEVICE;   // Hardware identifier
      Event_Class : Byte;   // Event class
      Fault_ID : Byte;   // Fault identifier
   END_VAR
BEGIN
END_ORGANIZATION_BLOCK

FUNCTION "Bypass assignments_0" : Void   // FC34, F_LAD
{ S7_Optimized_Access := 'TRUE' }
VERSION : 0.1
// stored: AutoNumber true, IsIECCheckEnabled false, UDAEnableTagReadback false
BEGIN

REGION Network 1
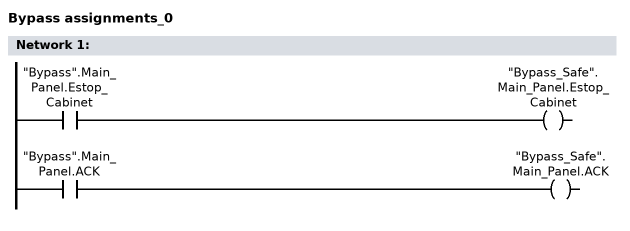
   RUNG wire#powerrail
      Contact( "Bypass".Main_Panel.Estop_Cabinet )
      Coil( "Bypass_Safe".Main_Panel.Estop_Cabinet )
   END_RUNG
   RUNG wire#powerrail
      Contact( "Bypass".Main_Panel.ACK )
      Coil( "Bypass_Safe".Main_Panel.ACK )
   END_RUNG
   // the same network as SCL:
   "Bypass_Safe".Main_Panel.Estop_Cabinet := "Bypass".Main_Panel.Estop_Cabinet;
   "Bypass_Safe".Main_Panel.ACK := "Bypass".Main_Panel.ACK;
END_REGION
END_FUNCTION

FUNCTION "Bypass assignments_1" : Void   // FC35, F_LAD
{ S7_Optimized_Access := 'TRUE' }
VERSION : 0.1
// stored: AutoNumber true, IsIECCheckEnabled false, UDAEnableTagReadback false
BEGIN

REGION Network 1
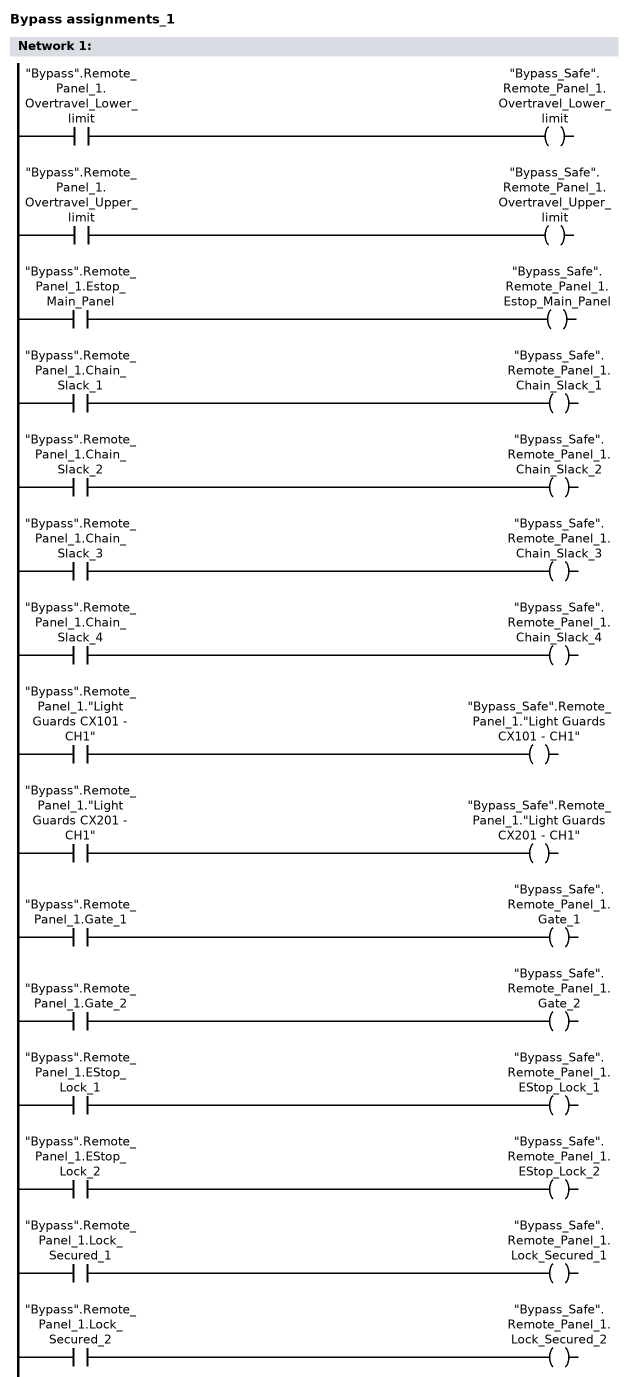
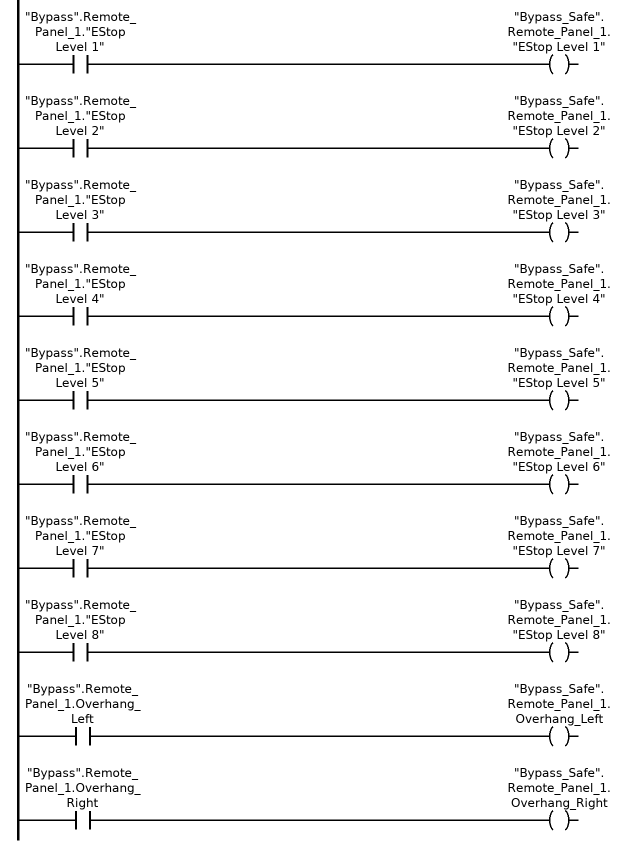
   RUNG wire#powerrail
      Contact( "Bypass".Remote_Panel_1.Overtravel_Lower_limit )
      Coil( "Bypass_Safe".Remote_Panel_1.Overtravel_Lower_limit )
   END_RUNG
   RUNG wire#powerrail
      Contact( "Bypass".Remote_Panel_1.Overtravel_Upper_limit )
      Coil( "Bypass_Safe".Remote_Panel_1.Overtravel_Upper_limit )
   END_RUNG
   RUNG wire#powerrail
      Contact( "Bypass".Remote_Panel_1.Estop_Main_Panel )
      Coil( "Bypass_Safe".Remote_Panel_1.Estop_Main_Panel )
   END_RUNG
   RUNG wire#powerrail
      Contact( "Bypass".Remote_Panel_1.Chain_Slack_1 )
      Coil( "Bypass_Safe".Remote_Panel_1.Chain_Slack_1 )
   END_RUNG
   RUNG wire#powerrail
      Contact( "Bypass".Remote_Panel_1.Chain_Slack_2 )
      Coil( "Bypass_Safe".Remote_Panel_1.Chain_Slack_2 )
   END_RUNG
   RUNG wire#powerrail
      Contact( "Bypass".Remote_Panel_1.Chain_Slack_3 )
      Coil( "Bypass_Safe".Remote_Panel_1.Chain_Slack_3 )
   END_RUNG
   RUNG wire#powerrail
      Contact( "Bypass".Remote_Panel_1.Chain_Slack_4 )
      Coil( "Bypass_Safe".Remote_Panel_1.Chain_Slack_4 )
   END_RUNG
   RUNG wire#powerrail
      Contact( "Bypass".Remote_Panel_1."Light Guards CX101 - CH1" )
      Coil( "Bypass_Safe".Remote_Panel_1."Light Guards CX101 - CH1" )
   END_RUNG
   RUNG wire#powerrail
      Contact( "Bypass".Remote_Panel_1."Light Guards CX201 - CH1" )
      Coil( "Bypass_Safe".Remote_Panel_1."Light Guards CX201 - CH1" )
   END_RUNG
   RUNG wire#powerrail
      Contact( "Bypass".Remote_Panel_1.Gate_1 )
      Coil( "Bypass_Safe".Remote_Panel_1.Gate_1 )
   END_RUNG
   RUNG wire#powerrail
      Contact( "Bypass".Remote_Panel_1.Gate_2 )
      Coil( "Bypass_Safe".Remote_Panel_1.Gate_2 )
   END_RUNG
   RUNG wire#powerrail
      Contact( "Bypass".Remote_Panel_1.EStop_Lock_1 )
      Coil( "Bypass_Safe".Remote_Panel_1.EStop_Lock_1 )
   END_RUNG
   RUNG wire#powerrail
      Contact( "Bypass".Remote_Panel_1.EStop_Lock_2 )
      Coil( "Bypass_Safe".Remote_Panel_1.EStop_Lock_2 )
   END_RUNG
   RUNG wire#powerrail
      Contact( "Bypass".Remote_Panel_1.Lock_Secured_1 )
      Coil( "Bypass_Safe".Remote_Panel_1.Lock_Secured_1 )
   END_RUNG
   RUNG wire#powerrail
      Contact( "Bypass".Remote_Panel_1.Lock_Secured_2 )
      Coil( "Bypass_Safe".Remote_Panel_1.Lock_Secured_2 )
   END_RUNG
   RUNG wire#powerrail
      Contact( "Bypass".Remote_Panel_1."EStop Level 1" )
      Coil( "Bypass_Safe".Remote_Panel_1."EStop Level 1" )
   END_RUNG
   RUNG wire#powerrail
      Contact( "Bypass".Remote_Panel_1."EStop Level 2" )
      Coil( "Bypass_Safe".Remote_Panel_1."EStop Level 2" )
   END_RUNG
   RUNG wire#powerrail
      Contact( "Bypass".Remote_Panel_1."EStop Level 3" )
      Coil( "Bypass_Safe".Remote_Panel_1."EStop Level 3" )
   END_RUNG
   RUNG wire#powerrail
      Contact( "Bypass".Remote_Panel_1."EStop Level 4" )
      Coil( "Bypass_Safe".Remote_Panel_1."EStop Level 4" )
   END_RUNG
   RUNG wire#powerrail
      Contact( "Bypass".Remote_Panel_1."EStop Level 5" )
      Coil( "Bypass_Safe".Remote_Panel_1."EStop Level 5" )
   END_RUNG
   RUNG wire#powerrail
      Contact( "Bypass".Remote_Panel_1."EStop Level 6" )
      Coil( "Bypass_Safe".Remote_Panel_1."EStop Level 6" )
   END_RUNG
   RUNG wire#powerrail
      Contact( "Bypass".Remote_Panel_1."EStop Level 7" )
      Coil( "Bypass_Safe".Remote_Panel_1."EStop Level 7" )
   END_RUNG
   RUNG wire#powerrail
      Contact( "Bypass".Remote_Panel_1."EStop Level 8" )
      Coil( "Bypass_Safe".Remote_Panel_1."EStop Level 8" )
   END_RUNG
   RUNG wire#powerrail
      Contact( "Bypass".Remote_Panel_1.Overhang_Left )
      Coil( "Bypass_Safe".Remote_Panel_1.Overhang_Left )
   END_RUNG
   RUNG wire#powerrail
      Contact( "Bypass".Remote_Panel_1.Overhang_Right )
      Coil( "Bypass_Safe".Remote_Panel_1.Overhang_Right )
   END_RUNG
   // the same network as SCL:
   "Bypass_Safe".Remote_Panel_1.Overtravel_Lower_limit := "Bypass".Remote_Panel_1.Overtravel_Lower_limit;
   "Bypass_Safe".Remote_Panel_1.Overtravel_Upper_limit := "Bypass".Remote_Panel_1.Overtravel_Upper_limit;
   "Bypass_Safe".Remote_Panel_1.Estop_Main_Panel := "Bypass".Remote_Panel_1.Estop_Main_Panel;
   "Bypass_Safe".Remote_Panel_1.Chain_Slack_1 := "Bypass".Remote_Panel_1.Chain_Slack_1;
   "Bypass_Safe".Remote_Panel_1.Chain_Slack_2 := "Bypass".Remote_Panel_1.Chain_Slack_2;
   "Bypass_Safe".Remote_Panel_1.Chain_Slack_3 := "Bypass".Remote_Panel_1.Chain_Slack_3;
   "Bypass_Safe".Remote_Panel_1.Chain_Slack_4 := "Bypass".Remote_Panel_1.Chain_Slack_4;
   "Bypass_Safe".Remote_Panel_1."Light Guards CX101 - CH1" := "Bypass".Remote_Panel_1."Light Guards CX101 - CH1";
   "Bypass_Safe".Remote_Panel_1."Light Guards CX201 - CH1" := "Bypass".Remote_Panel_1."Light Guards CX201 - CH1";
   "Bypass_Safe".Remote_Panel_1.Gate_1 := "Bypass".Remote_Panel_1.Gate_1;
   "Bypass_Safe".Remote_Panel_1.Gate_2 := "Bypass".Remote_Panel_1.Gate_2;
   "Bypass_Safe".Remote_Panel_1.EStop_Lock_1 := "Bypass".Remote_Panel_1.EStop_Lock_1;
   "Bypass_Safe".Remote_Panel_1.EStop_Lock_2 := "Bypass".Remote_Panel_1.EStop_Lock_2;
   "Bypass_Safe".Remote_Panel_1.Lock_Secured_1 := "Bypass".Remote_Panel_1.Lock_Secured_1;
   "Bypass_Safe".Remote_Panel_1.Lock_Secured_2 := "Bypass".Remote_Panel_1.Lock_Secured_2;
   "Bypass_Safe".Remote_Panel_1."EStop Level 1" := "Bypass".Remote_Panel_1."EStop Level 1";
   "Bypass_Safe".Remote_Panel_1."EStop Level 2" := "Bypass".Remote_Panel_1."EStop Level 2";
   "Bypass_Safe".Remote_Panel_1."EStop Level 3" := "Bypass".Remote_Panel_1."EStop Level 3";
   "Bypass_Safe".Remote_Panel_1."EStop Level 4" := "Bypass".Remote_Panel_1."EStop Level 4";
   "Bypass_Safe".Remote_Panel_1."EStop Level 5" := "Bypass".Remote_Panel_1."EStop Level 5";
   "Bypass_Safe".Remote_Panel_1."EStop Level 6" := "Bypass".Remote_Panel_1."EStop Level 6";
   "Bypass_Safe".Remote_Panel_1."EStop Level 7" := "Bypass".Remote_Panel_1."EStop Level 7";
   "Bypass_Safe".Remote_Panel_1."EStop Level 8" := "Bypass".Remote_Panel_1."EStop Level 8";
   "Bypass_Safe".Remote_Panel_1.Overhang_Left := "Bypass".Remote_Panel_1.Overhang_Left;
   "Bypass_Safe".Remote_Panel_1.Overhang_Right := "Bypass".Remote_Panel_1.Overhang_Right;
END_REGION
END_FUNCTION

FUNCTION "Bypass assignments_2" : Void   // FC36, F_LAD
{ S7_Optimized_Access := 'TRUE' }
VERSION : 0.1
// stored: AutoNumber true, IsIECCheckEnabled false, UDAEnableTagReadback false
BEGIN

REGION Network 1
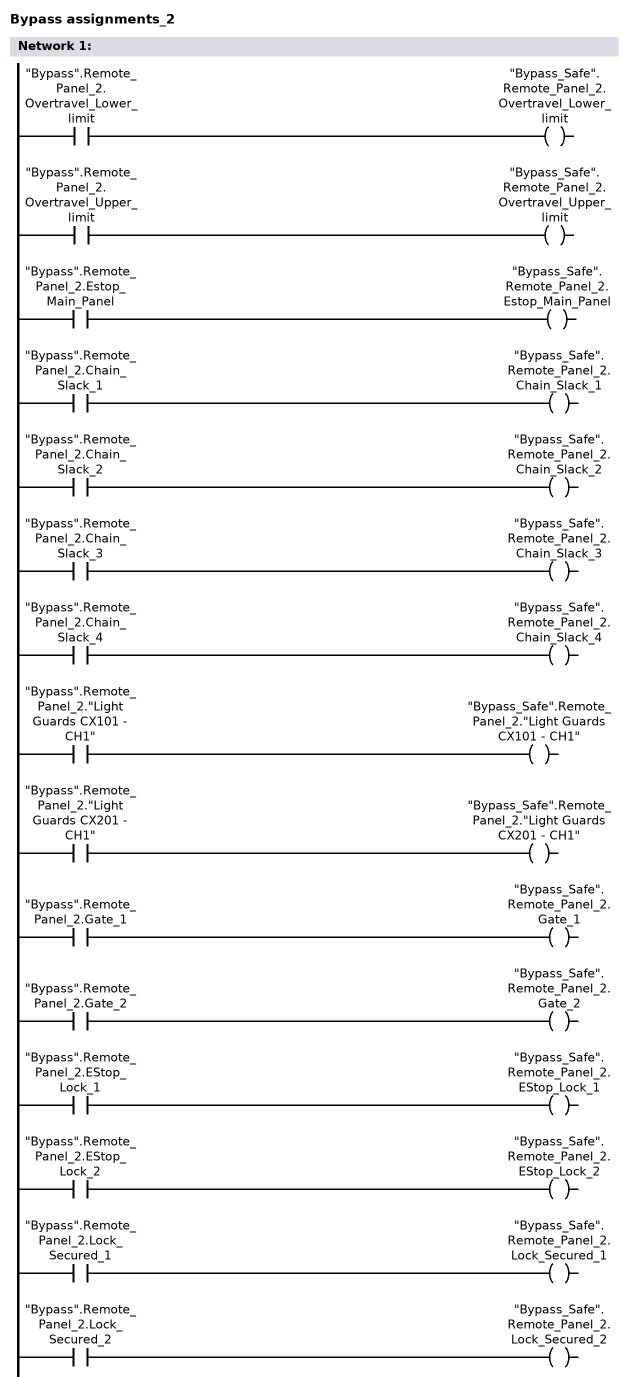
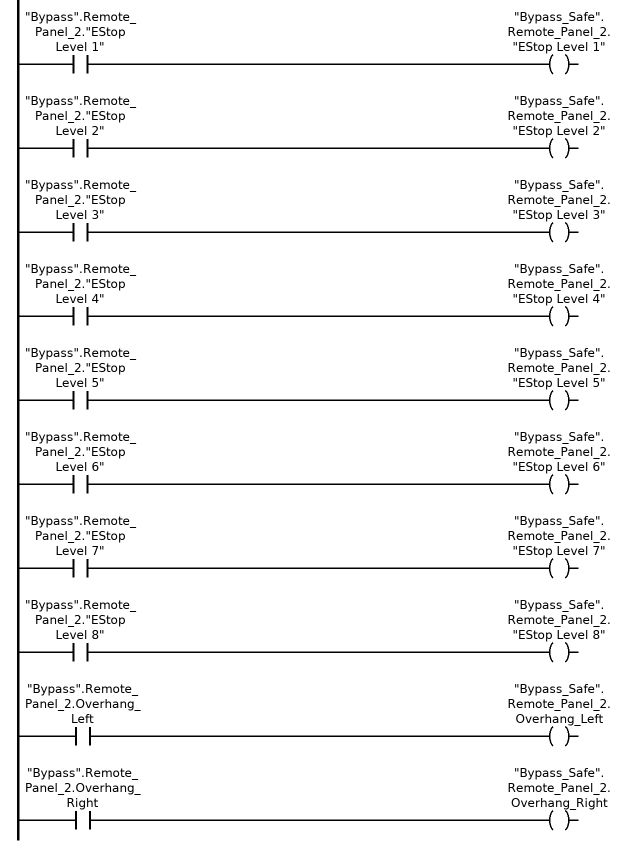
   RUNG wire#powerrail
      Contact( "Bypass".Remote_Panel_2.Overtravel_Lower_limit )
      Coil( "Bypass_Safe".Remote_Panel_2.Overtravel_Lower_limit )
   END_RUNG
   RUNG wire#powerrail
      Contact( "Bypass".Remote_Panel_2.Overtravel_Upper_limit )
      Coil( "Bypass_Safe".Remote_Panel_2.Overtravel_Upper_limit )
   END_RUNG
   RUNG wire#powerrail
      Contact( "Bypass".Remote_Panel_2.Estop_Main_Panel )
      Coil( "Bypass_Safe".Remote_Panel_2.Estop_Main_Panel )
   END_RUNG
   RUNG wire#powerrail
      Contact( "Bypass".Remote_Panel_2.Chain_Slack_1 )
      Coil( "Bypass_Safe".Remote_Panel_2.Chain_Slack_1 )
   END_RUNG
   RUNG wire#powerrail
      Contact( "Bypass".Remote_Panel_2.Chain_Slack_2 )
      Coil( "Bypass_Safe".Remote_Panel_2.Chain_Slack_2 )
   END_RUNG
   RUNG wire#powerrail
      Contact( "Bypass".Remote_Panel_2.Chain_Slack_3 )
      Coil( "Bypass_Safe".Remote_Panel_2.Chain_Slack_3 )
   END_RUNG
   RUNG wire#powerrail
      Contact( "Bypass".Remote_Panel_2.Chain_Slack_4 )
      Coil( "Bypass_Safe".Remote_Panel_2.Chain_Slack_4 )
   END_RUNG
   RUNG wire#powerrail
      Contact( "Bypass".Remote_Panel_2."Light Guards CX101 - CH1" )
      Coil( "Bypass_Safe".Remote_Panel_2."Light Guards CX101 - CH1" )
   END_RUNG
   RUNG wire#powerrail
      Contact( "Bypass".Remote_Panel_2."Light Guards CX201 - CH1" )
      Coil( "Bypass_Safe".Remote_Panel_2."Light Guards CX201 - CH1" )
   END_RUNG
   RUNG wire#powerrail
      Contact( "Bypass".Remote_Panel_2.Gate_1 )
      Coil( "Bypass_Safe".Remote_Panel_2.Gate_1 )
   END_RUNG
   RUNG wire#powerrail
      Contact( "Bypass".Remote_Panel_2.Gate_2 )
      Coil( "Bypass_Safe".Remote_Panel_2.Gate_2 )
   END_RUNG
   RUNG wire#powerrail
      Contact( "Bypass".Remote_Panel_2.EStop_Lock_1 )
      Coil( "Bypass_Safe".Remote_Panel_2.EStop_Lock_1 )
   END_RUNG
   RUNG wire#powerrail
      Contact( "Bypass".Remote_Panel_2.EStop_Lock_2 )
      Coil( "Bypass_Safe".Remote_Panel_2.EStop_Lock_2 )
   END_RUNG
   RUNG wire#powerrail
      Contact( "Bypass".Remote_Panel_2.Lock_Secured_1 )
      Coil( "Bypass_Safe".Remote_Panel_2.Lock_Secured_1 )
   END_RUNG
   RUNG wire#powerrail
      Contact( "Bypass".Remote_Panel_2.Lock_Secured_2 )
      Coil( "Bypass_Safe".Remote_Panel_2.Lock_Secured_2 )
   END_RUNG
   RUNG wire#powerrail
      Contact( "Bypass".Remote_Panel_2."EStop Level 1" )
      Coil( "Bypass_Safe".Remote_Panel_2."EStop Level 1" )
   END_RUNG
   RUNG wire#powerrail
      Contact( "Bypass".Remote_Panel_2."EStop Level 2" )
      Coil( "Bypass_Safe".Remote_Panel_2."EStop Level 2" )
   END_RUNG
   RUNG wire#powerrail
      Contact( "Bypass".Remote_Panel_2."EStop Level 3" )
      Coil( "Bypass_Safe".Remote_Panel_2."EStop Level 3" )
   END_RUNG
   RUNG wire#powerrail
      Contact( "Bypass".Remote_Panel_2."EStop Level 4" )
      Coil( "Bypass_Safe".Remote_Panel_2."EStop Level 4" )
   END_RUNG
   RUNG wire#powerrail
      Contact( "Bypass".Remote_Panel_2."EStop Level 5" )
      Coil( "Bypass_Safe".Remote_Panel_2."EStop Level 5" )
   END_RUNG
   RUNG wire#powerrail
      Contact( "Bypass".Remote_Panel_2."EStop Level 6" )
      Coil( "Bypass_Safe".Remote_Panel_2."EStop Level 6" )
   END_RUNG
   RUNG wire#powerrail
      Contact( "Bypass".Remote_Panel_2."EStop Level 7" )
      Coil( "Bypass_Safe".Remote_Panel_2."EStop Level 7" )
   END_RUNG
   RUNG wire#powerrail
      Contact( "Bypass".Remote_Panel_2."EStop Level 8" )
      Coil( "Bypass_Safe".Remote_Panel_2."EStop Level 8" )
   END_RUNG
   RUNG wire#powerrail
      Contact( "Bypass".Remote_Panel_2.Overhang_Left )
      Coil( "Bypass_Safe".Remote_Panel_2.Overhang_Left )
   END_RUNG
   RUNG wire#powerrail
      Contact( "Bypass".Remote_Panel_2.Overhang_Right )
      Coil( "Bypass_Safe".Remote_Panel_2.Overhang_Right )
   END_RUNG
   // the same network as SCL:
   "Bypass_Safe".Remote_Panel_2.Overtravel_Lower_limit := "Bypass".Remote_Panel_2.Overtravel_Lower_limit;
   "Bypass_Safe".Remote_Panel_2.Overtravel_Upper_limit := "Bypass".Remote_Panel_2.Overtravel_Upper_limit;
   "Bypass_Safe".Remote_Panel_2.Estop_Main_Panel := "Bypass".Remote_Panel_2.Estop_Main_Panel;
   "Bypass_Safe".Remote_Panel_2.Chain_Slack_1 := "Bypass".Remote_Panel_2.Chain_Slack_1;
   "Bypass_Safe".Remote_Panel_2.Chain_Slack_2 := "Bypass".Remote_Panel_2.Chain_Slack_2;
   "Bypass_Safe".Remote_Panel_2.Chain_Slack_3 := "Bypass".Remote_Panel_2.Chain_Slack_3;
   "Bypass_Safe".Remote_Panel_2.Chain_Slack_4 := "Bypass".Remote_Panel_2.Chain_Slack_4;
   "Bypass_Safe".Remote_Panel_2."Light Guards CX101 - CH1" := "Bypass".Remote_Panel_2."Light Guards CX101 - CH1";
   "Bypass_Safe".Remote_Panel_2."Light Guards CX201 - CH1" := "Bypass".Remote_Panel_2."Light Guards CX201 - CH1";
   "Bypass_Safe".Remote_Panel_2.Gate_1 := "Bypass".Remote_Panel_2.Gate_1;
   "Bypass_Safe".Remote_Panel_2.Gate_2 := "Bypass".Remote_Panel_2.Gate_2;
   "Bypass_Safe".Remote_Panel_2.EStop_Lock_1 := "Bypass".Remote_Panel_2.EStop_Lock_1;
   "Bypass_Safe".Remote_Panel_2.EStop_Lock_2 := "Bypass".Remote_Panel_2.EStop_Lock_2;
   "Bypass_Safe".Remote_Panel_2.Lock_Secured_1 := "Bypass".Remote_Panel_2.Lock_Secured_1;
   "Bypass_Safe".Remote_Panel_2.Lock_Secured_2 := "Bypass".Remote_Panel_2.Lock_Secured_2;
   "Bypass_Safe".Remote_Panel_2."EStop Level 1" := "Bypass".Remote_Panel_2."EStop Level 1";
   "Bypass_Safe".Remote_Panel_2."EStop Level 2" := "Bypass".Remote_Panel_2."EStop Level 2";
   "Bypass_Safe".Remote_Panel_2."EStop Level 3" := "Bypass".Remote_Panel_2."EStop Level 3";
   "Bypass_Safe".Remote_Panel_2."EStop Level 4" := "Bypass".Remote_Panel_2."EStop Level 4";
   "Bypass_Safe".Remote_Panel_2."EStop Level 5" := "Bypass".Remote_Panel_2."EStop Level 5";
   "Bypass_Safe".Remote_Panel_2."EStop Level 6" := "Bypass".Remote_Panel_2."EStop Level 6";
   "Bypass_Safe".Remote_Panel_2."EStop Level 7" := "Bypass".Remote_Panel_2."EStop Level 7";
   "Bypass_Safe".Remote_Panel_2."EStop Level 8" := "Bypass".Remote_Panel_2."EStop Level 8";
   "Bypass_Safe".Remote_Panel_2.Overhang_Left := "Bypass".Remote_Panel_2.Overhang_Left;
   "Bypass_Safe".Remote_Panel_2.Overhang_Right := "Bypass".Remote_Panel_2.Overhang_Right;
END_REGION
END_FUNCTION

FUNCTION "Bypass assignments_3" : Void   // FC37, F_LAD
{ S7_Optimized_Access := 'TRUE' }
VERSION : 0.1
// stored: AutoNumber true, IsIECCheckEnabled false, UDAEnableTagReadback false
BEGIN

REGION Network 1
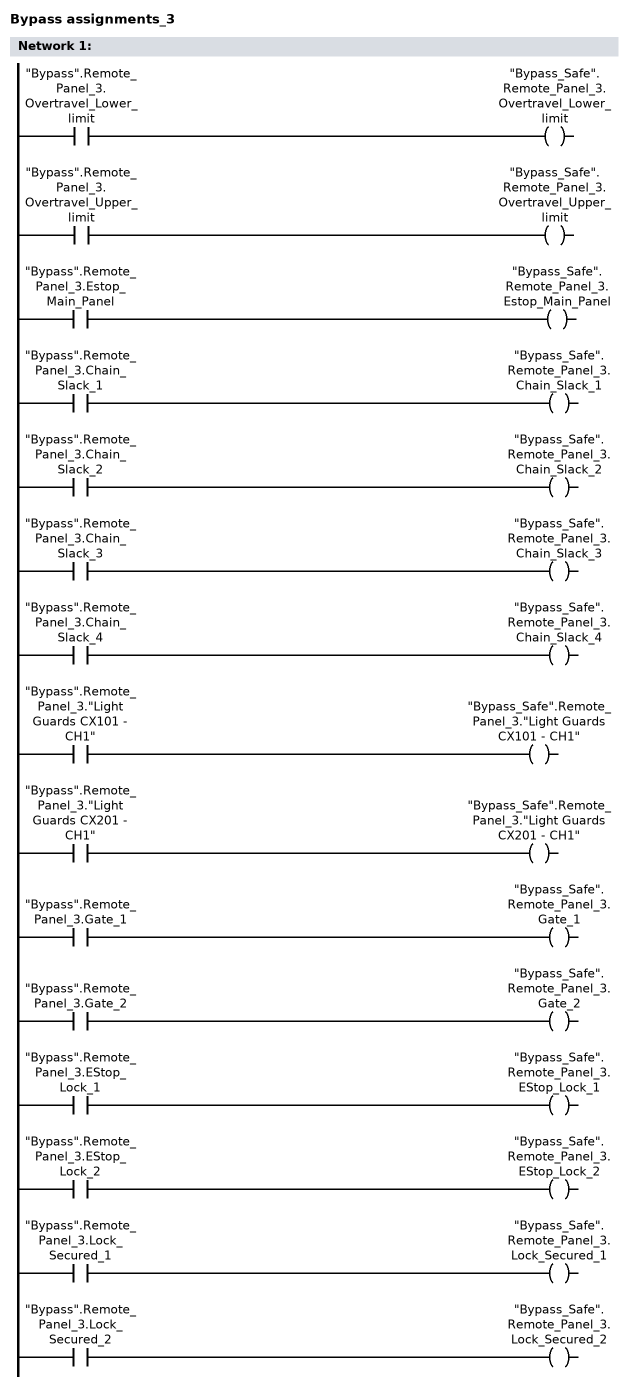
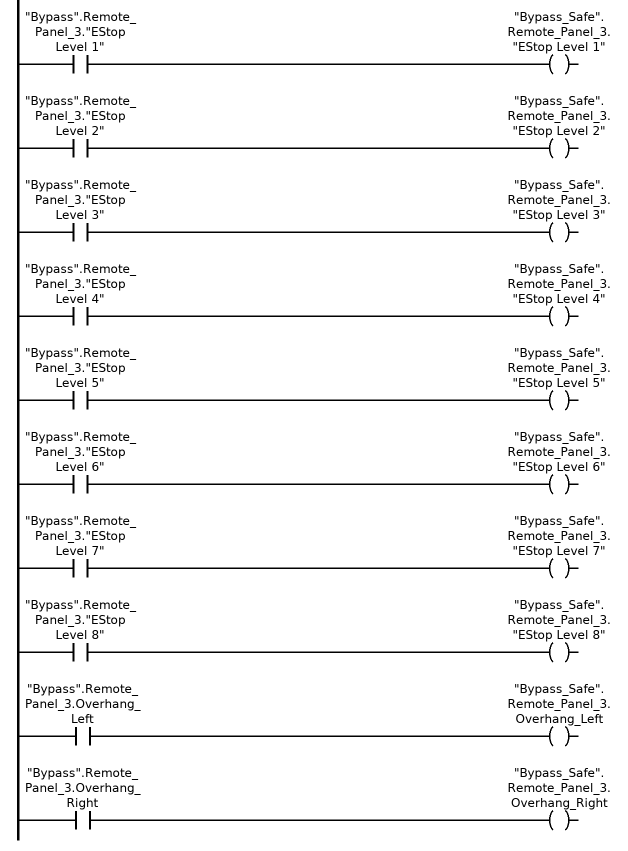
   RUNG wire#powerrail
      Contact( "Bypass".Remote_Panel_3.Overtravel_Lower_limit )
      Coil( "Bypass_Safe".Remote_Panel_3.Overtravel_Lower_limit )
   END_RUNG
   RUNG wire#powerrail
      Contact( "Bypass".Remote_Panel_3.Overtravel_Upper_limit )
      Coil( "Bypass_Safe".Remote_Panel_3.Overtravel_Upper_limit )
   END_RUNG
   RUNG wire#powerrail
      Contact( "Bypass".Remote_Panel_3.Estop_Main_Panel )
      Coil( "Bypass_Safe".Remote_Panel_3.Estop_Main_Panel )
   END_RUNG
   RUNG wire#powerrail
      Contact( "Bypass".Remote_Panel_3.Chain_Slack_1 )
      Coil( "Bypass_Safe".Remote_Panel_3.Chain_Slack_1 )
   END_RUNG
   RUNG wire#powerrail
      Contact( "Bypass".Remote_Panel_3.Chain_Slack_2 )
      Coil( "Bypass_Safe".Remote_Panel_3.Chain_Slack_2 )
   END_RUNG
   RUNG wire#powerrail
      Contact( "Bypass".Remote_Panel_3.Chain_Slack_3 )
      Coil( "Bypass_Safe".Remote_Panel_3.Chain_Slack_3 )
   END_RUNG
   RUNG wire#powerrail
      Contact( "Bypass".Remote_Panel_3.Chain_Slack_4 )
      Coil( "Bypass_Safe".Remote_Panel_3.Chain_Slack_4 )
   END_RUNG
   RUNG wire#powerrail
      Contact( "Bypass".Remote_Panel_3."Light Guards CX101 - CH1" )
      Coil( "Bypass_Safe".Remote_Panel_3."Light Guards CX101 - CH1" )
   END_RUNG
   RUNG wire#powerrail
      Contact( "Bypass".Remote_Panel_3."Light Guards CX201 - CH1" )
      Coil( "Bypass_Safe".Remote_Panel_3."Light Guards CX201 - CH1" )
   END_RUNG
   RUNG wire#powerrail
      Contact( "Bypass".Remote_Panel_3.Gate_1 )
      Coil( "Bypass_Safe".Remote_Panel_3.Gate_1 )
   END_RUNG
   RUNG wire#powerrail
      Contact( "Bypass".Remote_Panel_3.Gate_2 )
      Coil( "Bypass_Safe".Remote_Panel_3.Gate_2 )
   END_RUNG
   RUNG wire#powerrail
      Contact( "Bypass".Remote_Panel_3.EStop_Lock_1 )
      Coil( "Bypass_Safe".Remote_Panel_3.EStop_Lock_1 )
   END_RUNG
   RUNG wire#powerrail
      Contact( "Bypass".Remote_Panel_3.EStop_Lock_2 )
      Coil( "Bypass_Safe".Remote_Panel_3.EStop_Lock_2 )
   END_RUNG
   RUNG wire#powerrail
      Contact( "Bypass".Remote_Panel_3.Lock_Secured_1 )
      Coil( "Bypass_Safe".Remote_Panel_3.Lock_Secured_1 )
   END_RUNG
   RUNG wire#powerrail
      Contact( "Bypass".Remote_Panel_3.Lock_Secured_2 )
      Coil( "Bypass_Safe".Remote_Panel_3.Lock_Secured_2 )
   END_RUNG
   RUNG wire#powerrail
      Contact( "Bypass".Remote_Panel_3."EStop Level 1" )
      Coil( "Bypass_Safe".Remote_Panel_3."EStop Level 1" )
   END_RUNG
   RUNG wire#powerrail
      Contact( "Bypass".Remote_Panel_3."EStop Level 2" )
      Coil( "Bypass_Safe".Remote_Panel_3."EStop Level 2" )
   END_RUNG
   RUNG wire#powerrail
      Contact( "Bypass".Remote_Panel_3."EStop Level 3" )
      Coil( "Bypass_Safe".Remote_Panel_3."EStop Level 3" )
   END_RUNG
   RUNG wire#powerrail
      Contact( "Bypass".Remote_Panel_3."EStop Level 4" )
      Coil( "Bypass_Safe".Remote_Panel_3."EStop Level 4" )
   END_RUNG
   RUNG wire#powerrail
      Contact( "Bypass".Remote_Panel_3."EStop Level 5" )
      Coil( "Bypass_Safe".Remote_Panel_3."EStop Level 5" )
   END_RUNG
   RUNG wire#powerrail
      Contact( "Bypass".Remote_Panel_3."EStop Level 6" )
      Coil( "Bypass_Safe".Remote_Panel_3."EStop Level 6" )
   END_RUNG
   RUNG wire#powerrail
      Contact( "Bypass".Remote_Panel_3."EStop Level 7" )
      Coil( "Bypass_Safe".Remote_Panel_3."EStop Level 7" )
   END_RUNG
   RUNG wire#powerrail
      Contact( "Bypass".Remote_Panel_3."EStop Level 8" )
      Coil( "Bypass_Safe".Remote_Panel_3."EStop Level 8" )
   END_RUNG
   RUNG wire#powerrail
      Contact( "Bypass".Remote_Panel_3.Overhang_Left )
      Coil( "Bypass_Safe".Remote_Panel_3.Overhang_Left )
   END_RUNG
   RUNG wire#powerrail
      Contact( "Bypass".Remote_Panel_3.Overhang_Right )
      Coil( "Bypass_Safe".Remote_Panel_3.Overhang_Right )
   END_RUNG
   // the same network as SCL:
   "Bypass_Safe".Remote_Panel_3.Overtravel_Lower_limit := "Bypass".Remote_Panel_3.Overtravel_Lower_limit;
   "Bypass_Safe".Remote_Panel_3.Overtravel_Upper_limit := "Bypass".Remote_Panel_3.Overtravel_Upper_limit;
   "Bypass_Safe".Remote_Panel_3.Estop_Main_Panel := "Bypass".Remote_Panel_3.Estop_Main_Panel;
   "Bypass_Safe".Remote_Panel_3.Chain_Slack_1 := "Bypass".Remote_Panel_3.Chain_Slack_1;
   "Bypass_Safe".Remote_Panel_3.Chain_Slack_2 := "Bypass".Remote_Panel_3.Chain_Slack_2;
   "Bypass_Safe".Remote_Panel_3.Chain_Slack_3 := "Bypass".Remote_Panel_3.Chain_Slack_3;
   "Bypass_Safe".Remote_Panel_3.Chain_Slack_4 := "Bypass".Remote_Panel_3.Chain_Slack_4;
   "Bypass_Safe".Remote_Panel_3."Light Guards CX101 - CH1" := "Bypass".Remote_Panel_3."Light Guards CX101 - CH1";
   "Bypass_Safe".Remote_Panel_3."Light Guards CX201 - CH1" := "Bypass".Remote_Panel_3."Light Guards CX201 - CH1";
   "Bypass_Safe".Remote_Panel_3.Gate_1 := "Bypass".Remote_Panel_3.Gate_1;
   "Bypass_Safe".Remote_Panel_3.Gate_2 := "Bypass".Remote_Panel_3.Gate_2;
   "Bypass_Safe".Remote_Panel_3.EStop_Lock_1 := "Bypass".Remote_Panel_3.EStop_Lock_1;
   "Bypass_Safe".Remote_Panel_3.EStop_Lock_2 := "Bypass".Remote_Panel_3.EStop_Lock_2;
   "Bypass_Safe".Remote_Panel_3.Lock_Secured_1 := "Bypass".Remote_Panel_3.Lock_Secured_1;
   "Bypass_Safe".Remote_Panel_3.Lock_Secured_2 := "Bypass".Remote_Panel_3.Lock_Secured_2;
   "Bypass_Safe".Remote_Panel_3."EStop Level 1" := "Bypass".Remote_Panel_3."EStop Level 1";
   "Bypass_Safe".Remote_Panel_3."EStop Level 2" := "Bypass".Remote_Panel_3."EStop Level 2";
   "Bypass_Safe".Remote_Panel_3."EStop Level 3" := "Bypass".Remote_Panel_3."EStop Level 3";
   "Bypass_Safe".Remote_Panel_3."EStop Level 4" := "Bypass".Remote_Panel_3."EStop Level 4";
   "Bypass_Safe".Remote_Panel_3."EStop Level 5" := "Bypass".Remote_Panel_3."EStop Level 5";
   "Bypass_Safe".Remote_Panel_3."EStop Level 6" := "Bypass".Remote_Panel_3."EStop Level 6";
   "Bypass_Safe".Remote_Panel_3."EStop Level 7" := "Bypass".Remote_Panel_3."EStop Level 7";
   "Bypass_Safe".Remote_Panel_3."EStop Level 8" := "Bypass".Remote_Panel_3."EStop Level 8";
   "Bypass_Safe".Remote_Panel_3.Overhang_Left := "Bypass".Remote_Panel_3.Overhang_Left;
   "Bypass_Safe".Remote_Panel_3.Overhang_Right := "Bypass".Remote_Panel_3.Overhang_Right;
END_REGION
END_FUNCTION

FUNCTION "Bypass assignments_4" : Void   // FC39, F_LAD
{ S7_Optimized_Access := 'TRUE' }
VERSION : 0.1
// stored: AutoNumber true, IsIECCheckEnabled false, UDAEnableTagReadback false
BEGIN

REGION Network 1
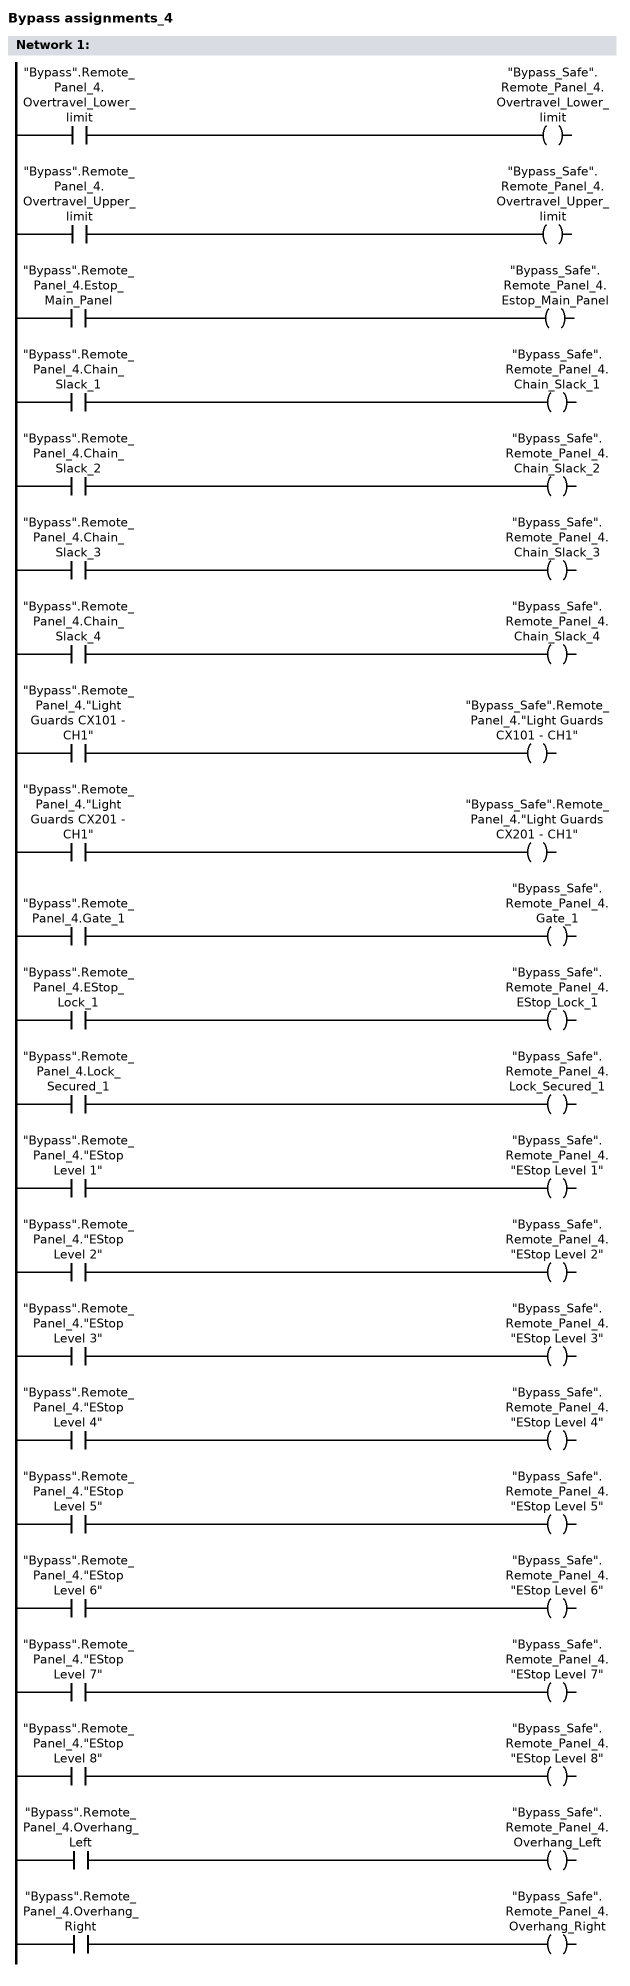
   RUNG wire#powerrail
      Contact( "Bypass".Remote_Panel_4.Overtravel_Lower_limit )
      Coil( "Bypass_Safe".Remote_Panel_4.Overtravel_Lower_limit )
   END_RUNG
   RUNG wire#powerrail
      Contact( "Bypass".Remote_Panel_4.Overtravel_Upper_limit )
      Coil( "Bypass_Safe".Remote_Panel_4.Overtravel_Upper_limit )
   END_RUNG
   RUNG wire#powerrail
      Contact( "Bypass".Remote_Panel_4.Estop_Main_Panel )
      Coil( "Bypass_Safe".Remote_Panel_4.Estop_Main_Panel )
   END_RUNG
   RUNG wire#powerrail
      Contact( "Bypass".Remote_Panel_4.Chain_Slack_1 )
      Coil( "Bypass_Safe".Remote_Panel_4.Chain_Slack_1 )
   END_RUNG
   RUNG wire#powerrail
      Contact( "Bypass".Remote_Panel_4.Chain_Slack_2 )
      Coil( "Bypass_Safe".Remote_Panel_4.Chain_Slack_2 )
   END_RUNG
   RUNG wire#powerrail
      Contact( "Bypass".Remote_Panel_4.Chain_Slack_3 )
      Coil( "Bypass_Safe".Remote_Panel_4.Chain_Slack_3 )
   END_RUNG
   RUNG wire#powerrail
      Contact( "Bypass".Remote_Panel_4.Chain_Slack_4 )
      Coil( "Bypass_Safe".Remote_Panel_4.Chain_Slack_4 )
   END_RUNG
   RUNG wire#powerrail
      Contact( "Bypass".Remote_Panel_4."Light Guards CX101 - CH1" )
      Coil( "Bypass_Safe".Remote_Panel_4."Light Guards CX101 - CH1" )
   END_RUNG
   RUNG wire#powerrail
      Contact( "Bypass".Remote_Panel_4."Light Guards CX201 - CH1" )
      Coil( "Bypass_Safe".Remote_Panel_4."Light Guards CX201 - CH1" )
   END_RUNG
   RUNG wire#powerrail
      Contact( "Bypass".Remote_Panel_4.Gate_1 )
      Coil( "Bypass_Safe".Remote_Panel_4.Gate_1 )
   END_RUNG
   RUNG wire#powerrail
      Contact( "Bypass".Remote_Panel_4.EStop_Lock_1 )
      Coil( "Bypass_Safe".Remote_Panel_4.EStop_Lock_1 )
   END_RUNG
   RUNG wire#powerrail
      Contact( "Bypass".Remote_Panel_4.Lock_Secured_1 )
      Coil( "Bypass_Safe".Remote_Panel_4.Lock_Secured_1 )
   END_RUNG
   RUNG wire#powerrail
      Contact( "Bypass".Remote_Panel_4."EStop Level 1" )
      Coil( "Bypass_Safe".Remote_Panel_4."EStop Level 1" )
   END_RUNG
   RUNG wire#powerrail
      Contact( "Bypass".Remote_Panel_4."EStop Level 2" )
      Coil( "Bypass_Safe".Remote_Panel_4."EStop Level 2" )
   END_RUNG
   RUNG wire#powerrail
      Contact( "Bypass".Remote_Panel_4."EStop Level 3" )
      Coil( "Bypass_Safe".Remote_Panel_4."EStop Level 3" )
   END_RUNG
   RUNG wire#powerrail
      Contact( "Bypass".Remote_Panel_4."EStop Level 4" )
      Coil( "Bypass_Safe".Remote_Panel_4."EStop Level 4" )
   END_RUNG
   RUNG wire#powerrail
      Contact( "Bypass".Remote_Panel_4."EStop Level 5" )
      Coil( "Bypass_Safe".Remote_Panel_4."EStop Level 5" )
   END_RUNG
   RUNG wire#powerrail
      Contact( "Bypass".Remote_Panel_4."EStop Level 6" )
      Coil( "Bypass_Safe".Remote_Panel_4."EStop Level 6" )
   END_RUNG
   RUNG wire#powerrail
      Contact( "Bypass".Remote_Panel_4."EStop Level 7" )
      Coil( "Bypass_Safe".Remote_Panel_4."EStop Level 7" )
   END_RUNG
   RUNG wire#powerrail
      Contact( "Bypass".Remote_Panel_4."EStop Level 8" )
      Coil( "Bypass_Safe".Remote_Panel_4."EStop Level 8" )
   END_RUNG
   RUNG wire#powerrail
      Contact( "Bypass".Remote_Panel_4.Overhang_Left )
      Coil( "Bypass_Safe".Remote_Panel_4.Overhang_Left )
   END_RUNG
   RUNG wire#powerrail
      Contact( "Bypass".Remote_Panel_4.Overhang_Right )
      Coil( "Bypass_Safe".Remote_Panel_4.Overhang_Right )
   END_RUNG
   // the same network as SCL:
   "Bypass_Safe".Remote_Panel_4.Overtravel_Lower_limit := "Bypass".Remote_Panel_4.Overtravel_Lower_limit;
   "Bypass_Safe".Remote_Panel_4.Overtravel_Upper_limit := "Bypass".Remote_Panel_4.Overtravel_Upper_limit;
   "Bypass_Safe".Remote_Panel_4.Estop_Main_Panel := "Bypass".Remote_Panel_4.Estop_Main_Panel;
   "Bypass_Safe".Remote_Panel_4.Chain_Slack_1 := "Bypass".Remote_Panel_4.Chain_Slack_1;
   "Bypass_Safe".Remote_Panel_4.Chain_Slack_2 := "Bypass".Remote_Panel_4.Chain_Slack_2;
   "Bypass_Safe".Remote_Panel_4.Chain_Slack_3 := "Bypass".Remote_Panel_4.Chain_Slack_3;
   "Bypass_Safe".Remote_Panel_4.Chain_Slack_4 := "Bypass".Remote_Panel_4.Chain_Slack_4;
   "Bypass_Safe".Remote_Panel_4."Light Guards CX101 - CH1" := "Bypass".Remote_Panel_4."Light Guards CX101 - CH1";
   "Bypass_Safe".Remote_Panel_4."Light Guards CX201 - CH1" := "Bypass".Remote_Panel_4."Light Guards CX201 - CH1";
   "Bypass_Safe".Remote_Panel_4.Gate_1 := "Bypass".Remote_Panel_4.Gate_1;
   "Bypass_Safe".Remote_Panel_4.EStop_Lock_1 := "Bypass".Remote_Panel_4.EStop_Lock_1;
   "Bypass_Safe".Remote_Panel_4.Lock_Secured_1 := "Bypass".Remote_Panel_4.Lock_Secured_1;
   "Bypass_Safe".Remote_Panel_4."EStop Level 1" := "Bypass".Remote_Panel_4."EStop Level 1";
   "Bypass_Safe".Remote_Panel_4."EStop Level 2" := "Bypass".Remote_Panel_4."EStop Level 2";
   "Bypass_Safe".Remote_Panel_4."EStop Level 3" := "Bypass".Remote_Panel_4."EStop Level 3";
   "Bypass_Safe".Remote_Panel_4."EStop Level 4" := "Bypass".Remote_Panel_4."EStop Level 4";
   "Bypass_Safe".Remote_Panel_4."EStop Level 5" := "Bypass".Remote_Panel_4."EStop Level 5";
   "Bypass_Safe".Remote_Panel_4."EStop Level 6" := "Bypass".Remote_Panel_4."EStop Level 6";
   "Bypass_Safe".Remote_Panel_4."EStop Level 7" := "Bypass".Remote_Panel_4."EStop Level 7";
   "Bypass_Safe".Remote_Panel_4."EStop Level 8" := "Bypass".Remote_Panel_4."EStop Level 8";
   "Bypass_Safe".Remote_Panel_4.Overhang_Left := "Bypass".Remote_Panel_4.Overhang_Left;
   "Bypass_Safe".Remote_Panel_4.Overhang_Right := "Bypass".Remote_Panel_4.Overhang_Right;
END_REGION
END_FUNCTION

FUNCTION "Bypass assignments_5" : Void   // FC38, F_LAD
{ S7_Optimized_Access := 'TRUE' }
VERSION : 0.1
// stored: AutoNumber true, IsIECCheckEnabled false, UDAEnableTagReadback false
BEGIN

REGION Network 1
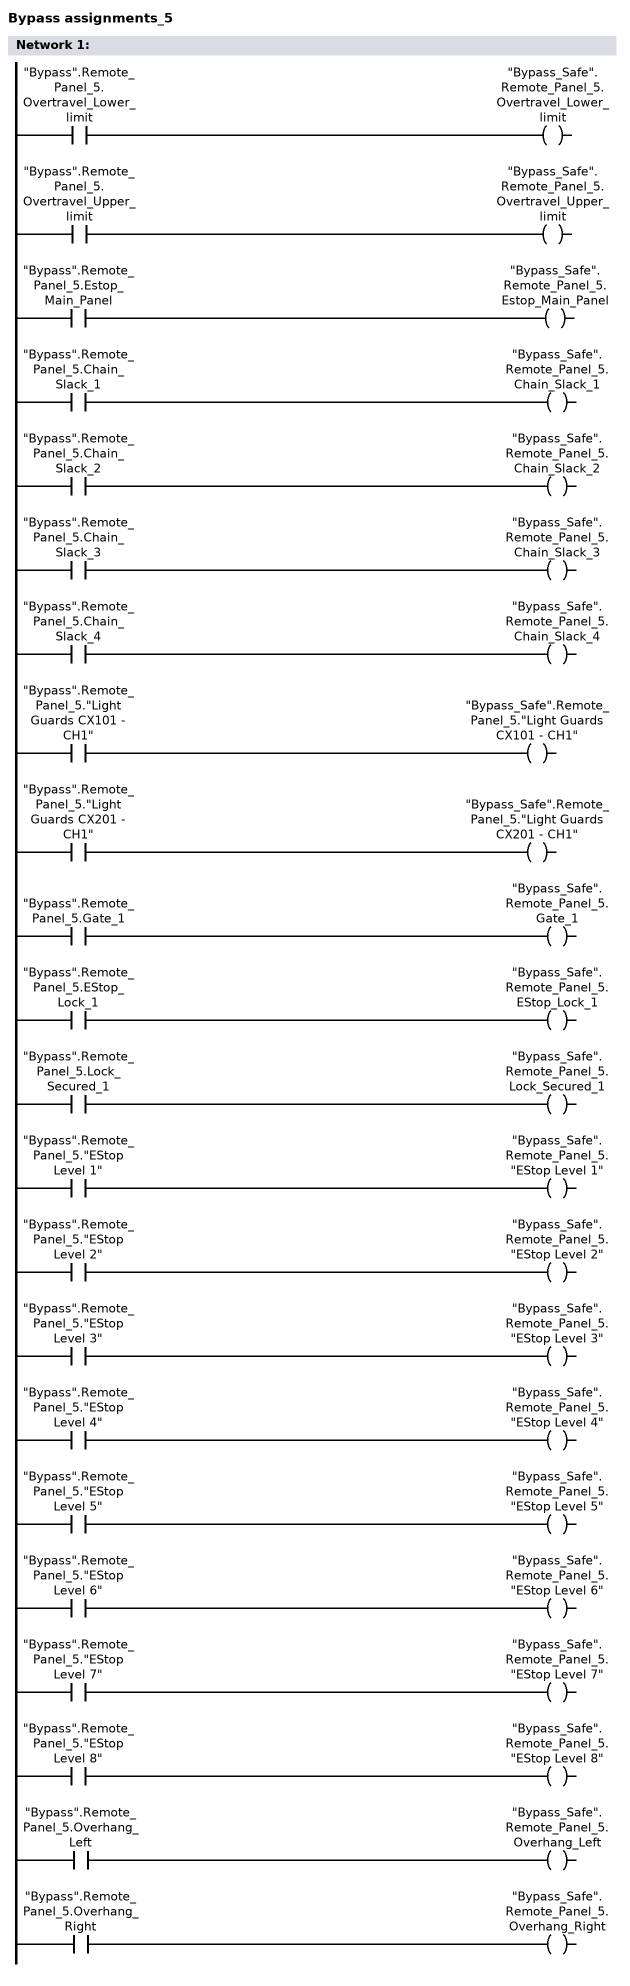
   RUNG wire#powerrail
      Contact( "Bypass".Remote_Panel_5.Overtravel_Lower_limit )
      Coil( "Bypass_Safe".Remote_Panel_5.Overtravel_Lower_limit )
   END_RUNG
   RUNG wire#powerrail
      Contact( "Bypass".Remote_Panel_5.Overtravel_Upper_limit )
      Coil( "Bypass_Safe".Remote_Panel_5.Overtravel_Upper_limit )
   END_RUNG
   RUNG wire#powerrail
      Contact( "Bypass".Remote_Panel_5.Estop_Main_Panel )
      Coil( "Bypass_Safe".Remote_Panel_5.Estop_Main_Panel )
   END_RUNG
   RUNG wire#powerrail
      Contact( "Bypass".Remote_Panel_5.Chain_Slack_1 )
      Coil( "Bypass_Safe".Remote_Panel_5.Chain_Slack_1 )
   END_RUNG
   RUNG wire#powerrail
      Contact( "Bypass".Remote_Panel_5.Chain_Slack_2 )
      Coil( "Bypass_Safe".Remote_Panel_5.Chain_Slack_2 )
   END_RUNG
   RUNG wire#powerrail
      Contact( "Bypass".Remote_Panel_5.Chain_Slack_3 )
      Coil( "Bypass_Safe".Remote_Panel_5.Chain_Slack_3 )
   END_RUNG
   RUNG wire#powerrail
      Contact( "Bypass".Remote_Panel_5.Chain_Slack_4 )
      Coil( "Bypass_Safe".Remote_Panel_5.Chain_Slack_4 )
   END_RUNG
   RUNG wire#powerrail
      Contact( "Bypass".Remote_Panel_5."Light Guards CX101 - CH1" )
      Coil( "Bypass_Safe".Remote_Panel_5."Light Guards CX101 - CH1" )
   END_RUNG
   RUNG wire#powerrail
      Contact( "Bypass".Remote_Panel_5."Light Guards CX201 - CH1" )
      Coil( "Bypass_Safe".Remote_Panel_5."Light Guards CX201 - CH1" )
   END_RUNG
   RUNG wire#powerrail
      Contact( "Bypass".Remote_Panel_5.Gate_1 )
      Coil( "Bypass_Safe".Remote_Panel_5.Gate_1 )
   END_RUNG
   RUNG wire#powerrail
      Contact( "Bypass".Remote_Panel_5.EStop_Lock_1 )
      Coil( "Bypass_Safe".Remote_Panel_5.EStop_Lock_1 )
   END_RUNG
   RUNG wire#powerrail
      Contact( "Bypass".Remote_Panel_5.Lock_Secured_1 )
      Coil( "Bypass_Safe".Remote_Panel_5.Lock_Secured_1 )
   END_RUNG
   RUNG wire#powerrail
      Contact( "Bypass".Remote_Panel_5."EStop Level 1" )
      Coil( "Bypass_Safe".Remote_Panel_5."EStop Level 1" )
   END_RUNG
   RUNG wire#powerrail
      Contact( "Bypass".Remote_Panel_5."EStop Level 2" )
      Coil( "Bypass_Safe".Remote_Panel_5."EStop Level 2" )
   END_RUNG
   RUNG wire#powerrail
      Contact( "Bypass".Remote_Panel_5."EStop Level 3" )
      Coil( "Bypass_Safe".Remote_Panel_5."EStop Level 3" )
   END_RUNG
   RUNG wire#powerrail
      Contact( "Bypass".Remote_Panel_5."EStop Level 4" )
      Coil( "Bypass_Safe".Remote_Panel_5."EStop Level 4" )
   END_RUNG
   RUNG wire#powerrail
      Contact( "Bypass".Remote_Panel_5."EStop Level 5" )
      Coil( "Bypass_Safe".Remote_Panel_5."EStop Level 5" )
   END_RUNG
   RUNG wire#powerrail
      Contact( "Bypass".Remote_Panel_5."EStop Level 6" )
      Coil( "Bypass_Safe".Remote_Panel_5."EStop Level 6" )
   END_RUNG
   RUNG wire#powerrail
      Contact( "Bypass".Remote_Panel_5."EStop Level 7" )
      Coil( "Bypass_Safe".Remote_Panel_5."EStop Level 7" )
   END_RUNG
   RUNG wire#powerrail
      Contact( "Bypass".Remote_Panel_5."EStop Level 8" )
      Coil( "Bypass_Safe".Remote_Panel_5."EStop Level 8" )
   END_RUNG
   RUNG wire#powerrail
      Contact( "Bypass".Remote_Panel_5.Overhang_Left )
      Coil( "Bypass_Safe".Remote_Panel_5.Overhang_Left )
   END_RUNG
   RUNG wire#powerrail
      Contact( "Bypass".Remote_Panel_5.Overhang_Right )
      Coil( "Bypass_Safe".Remote_Panel_5.Overhang_Right )
   END_RUNG
   // the same network as SCL:
   "Bypass_Safe".Remote_Panel_5.Overtravel_Lower_limit := "Bypass".Remote_Panel_5.Overtravel_Lower_limit;
   "Bypass_Safe".Remote_Panel_5.Overtravel_Upper_limit := "Bypass".Remote_Panel_5.Overtravel_Upper_limit;
   "Bypass_Safe".Remote_Panel_5.Estop_Main_Panel := "Bypass".Remote_Panel_5.Estop_Main_Panel;
   "Bypass_Safe".Remote_Panel_5.Chain_Slack_1 := "Bypass".Remote_Panel_5.Chain_Slack_1;
   "Bypass_Safe".Remote_Panel_5.Chain_Slack_2 := "Bypass".Remote_Panel_5.Chain_Slack_2;
   "Bypass_Safe".Remote_Panel_5.Chain_Slack_3 := "Bypass".Remote_Panel_5.Chain_Slack_3;
   "Bypass_Safe".Remote_Panel_5.Chain_Slack_4 := "Bypass".Remote_Panel_5.Chain_Slack_4;
   "Bypass_Safe".Remote_Panel_5."Light Guards CX101 - CH1" := "Bypass".Remote_Panel_5."Light Guards CX101 - CH1";
   "Bypass_Safe".Remote_Panel_5."Light Guards CX201 - CH1" := "Bypass".Remote_Panel_5."Light Guards CX201 - CH1";
   "Bypass_Safe".Remote_Panel_5.Gate_1 := "Bypass".Remote_Panel_5.Gate_1;
   "Bypass_Safe".Remote_Panel_5.EStop_Lock_1 := "Bypass".Remote_Panel_5.EStop_Lock_1;
   "Bypass_Safe".Remote_Panel_5.Lock_Secured_1 := "Bypass".Remote_Panel_5.Lock_Secured_1;
   "Bypass_Safe".Remote_Panel_5."EStop Level 1" := "Bypass".Remote_Panel_5."EStop Level 1";
   "Bypass_Safe".Remote_Panel_5."EStop Level 2" := "Bypass".Remote_Panel_5."EStop Level 2";
   "Bypass_Safe".Remote_Panel_5."EStop Level 3" := "Bypass".Remote_Panel_5."EStop Level 3";
   "Bypass_Safe".Remote_Panel_5."EStop Level 4" := "Bypass".Remote_Panel_5."EStop Level 4";
   "Bypass_Safe".Remote_Panel_5."EStop Level 5" := "Bypass".Remote_Panel_5."EStop Level 5";
   "Bypass_Safe".Remote_Panel_5."EStop Level 6" := "Bypass".Remote_Panel_5."EStop Level 6";
   "Bypass_Safe".Remote_Panel_5."EStop Level 7" := "Bypass".Remote_Panel_5."EStop Level 7";
   "Bypass_Safe".Remote_Panel_5."EStop Level 8" := "Bypass".Remote_Panel_5."EStop Level 8";
   "Bypass_Safe".Remote_Panel_5.Overhang_Left := "Bypass".Remote_Panel_5.Overhang_Left;
   "Bypass_Safe".Remote_Panel_5.Overhang_Right := "Bypass".Remote_Panel_5.Overhang_Right;
END_REGION
END_FUNCTION

FUNCTION "ByteArrayToString" : String   // FC15, SCL
{ S7_Optimized_Access := 'TRUE' }
VERSION : 0.1
// stored: AutoNumber true, IsIECCheckEnabled false, SetENOAutomatically false, UDAEnableTagReadback false
   VAR_INPUT
      Lenght : Int;
      ByteArray : Array[0..1024] of Byte;
   END_VAR
   VAR_OUTPUT
      ByteArrayToString_1 : String;
      ByteArrayToString_2 : String;
      ByteArrayToString_3 : String;
      ByteArrayToString_4 : String;
      ByteArrayToString_5 : String;
   END_VAR
   VAR_TEMP
      tempStr_1 : String;
      tempStr_2 : String;
      tempStr_3 : String;
      tempStr_4 : String;
      tempStr_5 : String;
      tempStr_6 : String;
      foundPos : Int;
      i : Int;
   END_VAR
BEGIN
   //STRING 1
   #tempStr_1 := '';
   FOR #i := 0 TO MIN(IN1 := #Lenght - 1, IN2 := 254) DO
       IF #ByteArray[#i] <> 0 THEN
           #tempStr_1 := CONCAT(IN1 := #tempStr_1, IN2 := CHAR_TO_STRING(BYTE_TO_CHAR(#ByteArray[#i])));
       END_IF;
   END_FOR;

   //STRING 2
   #tempStr_2 := '';
   FOR #i := 100 TO MIN(IN1 := #Lenght - 1, IN2 := 354) DO
       IF #ByteArray[#i] <> 0 THEN
           #tempStr_2 := CONCAT(IN1 := #tempStr_2, IN2 := CHAR_TO_STRING(BYTE_TO_CHAR(#ByteArray[#i])));
       END_IF;
   END_FOR;

   //STRING 3
   #tempStr_3 := '';
   FOR #i := 200 TO MIN(IN1 := #Lenght - 1, IN2 := 454) DO
       IF #ByteArray[#i] <> 0 THEN
           #tempStr_3 := CONCAT(IN1 := #tempStr_3, IN2 := CHAR_TO_STRING(BYTE_TO_CHAR(#ByteArray[#i])));
       END_IF;
   END_FOR;

   //STRING 4
   #tempStr_4 := '';
   FOR #i := 300 TO MIN(IN1 := #Lenght - 1, IN2 := 554) DO
       IF #ByteArray[#i] <> 0 THEN
           #tempStr_4 := CONCAT(IN1 := #tempStr_4, IN2 := CHAR_TO_STRING(BYTE_TO_CHAR(#ByteArray[#i])));
       END_IF;
   END_FOR;

   // //STRING 5
   #tempStr_5 := '';
   FOR #i := 400 TO MIN(IN1 := #Lenght - 1, IN2 := 654) DO
       IF #ByteArray[#i] <> 0 THEN
           #tempStr_5 := CONCAT(IN1 := #tempStr_5, IN2 := CHAR_TO_STRING(BYTE_TO_CHAR(#ByteArray[#i])));
       END_IF;
   END_FOR;

   // //STRING 6
   #tempStr_6 := '';
   FOR #i := 500 TO MIN(IN1 := #Lenght - 1, IN2 := 763) DO
       IF #ByteArray[#i] <> 0 THEN
           #tempStr_6 := CONCAT(IN1 := #tempStr_6, IN2 := CHAR_TO_STRING(BYTE_TO_CHAR(#ByteArray[#i])));
       END_IF;
   END_FOR;

   // Remove '$R$L'
   // string 1
   #foundPos := FIND(IN1 := #tempStr_1, IN2 := '$R$L');
   WHILE #foundPos > 0 DO
       #tempStr_1 := REPLACE(IN1 := #tempStr_1, IN2 := '', P := #foundPos, L := 2);
       #foundPos := FIND(IN1 := #tempStr_1, IN2 := '$R$L');
   END_WHILE;

   // string 2
   #foundPos := FIND(IN1 := #tempStr_2, IN2 := '$R$L');
   WHILE #foundPos > 0 DO
       #tempStr_2 := REPLACE(IN1 := #tempStr_2, IN2 := '', P := #foundPos, L := 2);
       #foundPos := FIND(IN1 := #tempStr_2, IN2 := '$R$L');
   END_WHILE;

   // string 3
   #foundPos := FIND(IN1 := #tempStr_3, IN2 := '$R$L');
   WHILE #foundPos > 0 DO
       #tempStr_3 := REPLACE(IN1 := #tempStr_3, IN2 := '', P := #foundPos, L := 2);
       #foundPos := FIND(IN1 := #tempStr_3, IN2 := '$R$L');
   END_WHILE;

   // string 4
   #foundPos := FIND(IN1 := #tempStr_4, IN2 := '$R$L');
   WHILE #foundPos > 0 DO
       #tempStr_4 := REPLACE(IN1 := #tempStr_4, IN2 := '', P := #foundPos, L := 2);
       #foundPos := FIND(IN1 := #tempStr_4, IN2 := '$R$L');
   END_WHILE;

   // string 5
   #foundPos := FIND(IN1 := #tempStr_5, IN2 := '$R$L');
   WHILE #foundPos > 0 DO
       #tempStr_5 := REPLACE(IN1 := #tempStr_5, IN2 := '', P := #foundPos, L := 2);
       #foundPos := FIND(IN1 := #tempStr_5, IN2 := '$R$L');
   END_WHILE;

   // string 6
   #foundPos := FIND(IN1 := #tempStr_6, IN2 := '$R$L');
   WHILE #foundPos > 0 DO
       #tempStr_6 := REPLACE(IN1 := #tempStr_6, IN2 := '', P := #foundPos, L := 2);
       #foundPos := FIND(IN1 := #tempStr_6, IN2 := '$R$L');
   END_WHILE;

   #ByteArrayToString := #tempStr_1;
   #ByteArrayToString_1 := #tempStr_2;
   #ByteArrayToString_2 := #tempStr_3;
   #ByteArrayToString_3 := #tempStr_4;
   #ByteArrayToString_4 := #tempStr_5;
   #ByteArrayToString_5 := #tempStr_6;
END_FUNCTION

FUNCTION "ByteArrayToString_1" : String   // FC23, SCL
{ S7_Optimized_Access := 'TRUE' }
VERSION : 0.1
// stored: AutoNumber true, IsIECCheckEnabled false, SetENOAutomatically false, UDAEnableTagReadback false
   VAR_INPUT
      Lenght : Int;
      ByteArray : Array[1..200] of Byte;
   END_VAR
   VAR_TEMP
      tempStr_1 : String;
      foundPos : Int;
      i : Int;
   END_VAR
BEGIN
   #tempStr_1 := '';
   FOR #i := 1 TO MIN(IN1 := #Lenght - 1, IN2 := 200) DO
       IF #ByteArray[#i] <> 0 THEN
           #tempStr_1 := CONCAT(IN1 := #tempStr_1, IN2 := CHAR_TO_STRING(BYTE_TO_CHAR(#ByteArray[#i])));
       END_IF;
   END_FOR;

   // Remove '$02'
   // string 1
   #foundPos := FIND(IN1 := #tempStr_1, IN2 := '$02');
   WHILE #foundPos > 0 DO
       #tempStr_1 := REPLACE(IN1 := #tempStr_1, IN2 := '', P := #foundPos, L := 1);
       #foundPos := FIND(IN1 := #tempStr_1, IN2 := '$02');
   END_WHILE;

   #ByteArrayToString_1 := #tempStr_1;
END_FUNCTION

FUNCTION "CNV_Charge_Settings_FC" : Void   // FC42, SCL
{ S7_Optimized_Access := 'TRUE' }
VERSION : 0.1
// stored: AutoNumber true, IsIECCheckEnabled false, SetENOAutomatically false, UDAEnableTagReadback false
BEGIN
   CASE "CNV_System_Selected" OF
       1: //SYSTEM 1
           CASE "CNV_Level_Selected" OF
               1:
                   "PopUps_DB".Buffer_Cnv_Settings_1 := "Settings_DB".LCnv_Sys[1].Cnv_Level[1].Cnv1;
                   "PopUps_DB".ECnv_Settings := "Settings_DB".ECnv_Sys[1];
                   "PopUps_DB".Buffer_Cnv_Settings_2 := "Settings_DB".LCnv_Sys[1].Cnv_Level[1].Cnv2;
               2:
                   "PopUps_DB".Buffer_Cnv_Settings_1 := "Settings_DB".LCnv_Sys[1].Cnv_Level[2].Cnv1;
                   "PopUps_DB".ECnv_Settings := "Settings_DB".ECnv_Sys[1];
                   "PopUps_DB".Buffer_Cnv_Settings_2 := "Settings_DB".LCnv_Sys[1].Cnv_Level[2].Cnv2;
               3:
                   "PopUps_DB".Buffer_Cnv_Settings_1 := "Settings_DB".LCnv_Sys[1].Cnv_Level[3].Cnv1;
                   "PopUps_DB".ECnv_Settings := "Settings_DB".ECnv_Sys[1];
                   "PopUps_DB".Buffer_Cnv_Settings_2 := "Settings_DB".LCnv_Sys[1].Cnv_Level[3].Cnv2;
               4:
                   "PopUps_DB".Buffer_Cnv_Settings_1 := "Settings_DB".LCnv_Sys[1].Cnv_Level[4].Cnv1;
                   "PopUps_DB".ECnv_Settings := "Settings_DB".ECnv_Sys[1];
                   "PopUps_DB".Buffer_Cnv_Settings_2 := "Settings_DB".LCnv_Sys[1].Cnv_Level[4].Cnv2;
               5:
                   "PopUps_DB".Buffer_Cnv_Settings_1 := "Settings_DB".LCnv_Sys[1].Cnv_Level[5].Cnv1;
                   "PopUps_DB".ECnv_Settings := "Settings_DB".ECnv_Sys[1];
                   "PopUps_DB".Buffer_Cnv_Settings_2 := "Settings_DB".LCnv_Sys[1].Cnv_Level[5].Cnv2;
               6:
                   "PopUps_DB".Buffer_Cnv_Settings_1 := "Settings_DB".LCnv_Sys[1].Cnv_Level[6].Cnv1;
                   "PopUps_DB".ECnv_Settings := "Settings_DB".ECnv_Sys[1];
                   "PopUps_DB".Buffer_Cnv_Settings_2 := "Settings_DB".LCnv_Sys[1].Cnv_Level[6].Cnv2;
               7:
                   "PopUps_DB".Buffer_Cnv_Settings_1 := "Settings_DB".LCnv_Sys[1].Cnv_Level[7].Cnv1;
                   "PopUps_DB".ECnv_Settings := "Settings_DB".ECnv_Sys[1];
                   "PopUps_DB".Buffer_Cnv_Settings_2 := "Settings_DB".LCnv_Sys[1].Cnv_Level[7].Cnv2;
               8:
                   "PopUps_DB".Buffer_Cnv_Settings_1 := "Settings_DB".LCnv_Sys[1].Cnv_Level[8].Cnv1;
                   "PopUps_DB".ECnv_Settings := "Settings_DB".ECnv_Sys[1];
                   "PopUps_DB".Buffer_Cnv_Settings_2 := "Settings_DB".LCnv_Sys[1].Cnv_Level[8].Cnv2;
           END_CASE;
       2: //SYSTEM 2
           CASE "CNV_Level_Selected" OF
               1:
                   "PopUps_DB".Buffer_Cnv_Settings_1 := "Settings_DB".LCnv_Sys[2].Cnv_Level[1].Cnv1;
                   "PopUps_DB".ECnv_Settings := "Settings_DB".ECnv_Sys[2];
                   "PopUps_DB".Buffer_Cnv_Settings_2 := "Settings_DB".LCnv_Sys[2].Cnv_Level[1].Cnv2;
               2:
                   "PopUps_DB".Buffer_Cnv_Settings_1 := "Settings_DB".LCnv_Sys[2].Cnv_Level[2].Cnv1;
                   "PopUps_DB".ECnv_Settings := "Settings_DB".ECnv_Sys[2];
                   "PopUps_DB".Buffer_Cnv_Settings_2 := "Settings_DB".LCnv_Sys[2].Cnv_Level[2].Cnv2;
               3:
                   "PopUps_DB".Buffer_Cnv_Settings_1 := "Settings_DB".LCnv_Sys[2].Cnv_Level[3].Cnv1;
                   "PopUps_DB".ECnv_Settings := "Settings_DB".ECnv_Sys[2];
                   "PopUps_DB".Buffer_Cnv_Settings_2 := "Settings_DB".LCnv_Sys[2].Cnv_Level[3].Cnv2;
               4:
                   "PopUps_DB".Buffer_Cnv_Settings_1 := "Settings_DB".LCnv_Sys[2].Cnv_Level[4].Cnv1;
                   "PopUps_DB".ECnv_Settings := "Settings_DB".ECnv_Sys[2];
                   "PopUps_DB".Buffer_Cnv_Settings_2 := "Settings_DB".LCnv_Sys[2].Cnv_Level[4].Cnv2;
               5:
                   "PopUps_DB".Buffer_Cnv_Settings_1 := "Settings_DB".LCnv_Sys[2].Cnv_Level[5].Cnv1;
                   "PopUps_DB".ECnv_Settings := "Settings_DB".ECnv_Sys[2];
                   "PopUps_DB".Buffer_Cnv_Settings_2 := "Settings_DB".LCnv_Sys[2].Cnv_Level[5].Cnv2;
               6:
                   "PopUps_DB".Buffer_Cnv_Settings_1 := "Settings_DB".LCnv_Sys[2].Cnv_Level[6].Cnv1;
                   "PopUps_DB".ECnv_Settings := "Settings_DB".ECnv_Sys[2];
                   "PopUps_DB".Buffer_Cnv_Settings_2 := "Settings_DB".LCnv_Sys[2].Cnv_Level[6].Cnv2;
               7:
                   "PopUps_DB".Buffer_Cnv_Settings_1 := "Settings_DB".LCnv_Sys[2].Cnv_Level[7].Cnv1;
                   "PopUps_DB".ECnv_Settings := "Settings_DB".ECnv_Sys[2];
                   "PopUps_DB".Buffer_Cnv_Settings_2 := "Settings_DB".LCnv_Sys[2].Cnv_Level[7].Cnv2;
               8:
                   "PopUps_DB".Buffer_Cnv_Settings_1 := "Settings_DB".LCnv_Sys[2].Cnv_Level[8].Cnv1;
                   "PopUps_DB".ECnv_Settings := "Settings_DB".ECnv_Sys[2];
                   "PopUps_DB".Buffer_Cnv_Settings_2 := "Settings_DB".LCnv_Sys[2].Cnv_Level[8].Cnv2;
           END_CASE;
       3: //SYSTEM 3
           CASE "CNV_Level_Selected" OF
               1:
                   "PopUps_DB".Buffer_Cnv_Settings_1 := "Settings_DB".LCnv_Sys[3].Cnv_Level[1].Cnv1;
                   "PopUps_DB".ECnv_Settings := "Settings_DB".ECnv_Sys[3];
                   "PopUps_DB".Buffer_Cnv_Settings_2 := "Settings_DB".LCnv_Sys[3].Cnv_Level[1].Cnv2;
               2:
                   "PopUps_DB".Buffer_Cnv_Settings_1 := "Settings_DB".LCnv_Sys[3].Cnv_Level[2].Cnv1;
                   "PopUps_DB".ECnv_Settings := "Settings_DB".ECnv_Sys[3];
                   "PopUps_DB".Buffer_Cnv_Settings_2 := "Settings_DB".LCnv_Sys[3].Cnv_Level[2].Cnv2;
               3:
                   "PopUps_DB".Buffer_Cnv_Settings_1 := "Settings_DB".LCnv_Sys[3].Cnv_Level[3].Cnv1;
                   "PopUps_DB".ECnv_Settings := "Settings_DB".ECnv_Sys[3];
                   "PopUps_DB".Buffer_Cnv_Settings_2 := "Settings_DB".LCnv_Sys[3].Cnv_Level[3].Cnv2;
               4:
                   "PopUps_DB".Buffer_Cnv_Settings_1 := "Settings_DB".LCnv_Sys[3].Cnv_Level[4].Cnv1;
                   "PopUps_DB".ECnv_Settings := "Settings_DB".ECnv_Sys[3];
                   "PopUps_DB".Buffer_Cnv_Settings_2 := "Settings_DB".LCnv_Sys[3].Cnv_Level[4].Cnv2;
               5:
                   "PopUps_DB".Buffer_Cnv_Settings_1 := "Settings_DB".LCnv_Sys[3].Cnv_Level[5].Cnv1;
                   "PopUps_DB".ECnv_Settings := "Settings_DB".ECnv_Sys[3];
                   "PopUps_DB".Buffer_Cnv_Settings_2 := "Settings_DB".LCnv_Sys[3].Cnv_Level[5].Cnv2;
               6:
                   "PopUps_DB".Buffer_Cnv_Settings_1 := "Settings_DB".LCnv_Sys[3].Cnv_Level[6].Cnv1;
                   "PopUps_DB".ECnv_Settings := "Settings_DB".ECnv_Sys[3];
                   "PopUps_DB".Buffer_Cnv_Settings_2 := "Settings_DB".LCnv_Sys[3].Cnv_Level[6].Cnv2;
               7:
                   "PopUps_DB".Buffer_Cnv_Settings_1 := "Settings_DB".LCnv_Sys[3].Cnv_Level[7].Cnv1;
                   "PopUps_DB".ECnv_Settings := "Settings_DB".ECnv_Sys[3];
                   "PopUps_DB".Buffer_Cnv_Settings_2 := "Settings_DB".LCnv_Sys[3].Cnv_Level[7].Cnv2;
               8:
                   "PopUps_DB".Buffer_Cnv_Settings_1 := "Settings_DB".LCnv_Sys[3].Cnv_Level[8].Cnv1;
                   "PopUps_DB".ECnv_Settings := "Settings_DB".ECnv_Sys[3];
                   "PopUps_DB".Buffer_Cnv_Settings_2 := "Settings_DB".LCnv_Sys[3].Cnv_Level[8].Cnv2;
           END_CASE;
       4: //SYSTEM 4
           CASE "CNV_Level_Selected" OF
               1:
                   "PopUps_DB".Buffer_Cnv_Settings_1 := "Settings_DB".LCnv_Sys[4].Cnv_Level[1].Cnv1;
                   "PopUps_DB".ECnv_Settings := "Settings_DB".ECnv_Sys[4];
                   "PopUps_DB".Buffer_Cnv_Settings_2 := "Settings_DB".LCnv_Sys[4].Cnv_Level[1].Cnv2;
               2:
                   "PopUps_DB".Buffer_Cnv_Settings_1 := "Settings_DB".LCnv_Sys[4].Cnv_Level[2].Cnv1;
                   "PopUps_DB".ECnv_Settings := "Settings_DB".ECnv_Sys[4];
                   "PopUps_DB".Buffer_Cnv_Settings_2 := "Settings_DB".LCnv_Sys[4].Cnv_Level[2].Cnv2;
               3:
                   "PopUps_DB".Buffer_Cnv_Settings_1 := "Settings_DB".LCnv_Sys[4].Cnv_Level[3].Cnv1;
                   "PopUps_DB".ECnv_Settings := "Settings_DB".ECnv_Sys[4];
                   "PopUps_DB".Buffer_Cnv_Settings_2 := "Settings_DB".LCnv_Sys[4].Cnv_Level[3].Cnv2;
               4:
                   "PopUps_DB".Buffer_Cnv_Settings_1 := "Settings_DB".LCnv_Sys[4].Cnv_Level[4].Cnv1;
                   "PopUps_DB".ECnv_Settings := "Settings_DB".ECnv_Sys[4];
                   "PopUps_DB".Buffer_Cnv_Settings_2 := "Settings_DB".LCnv_Sys[4].Cnv_Level[4].Cnv2;
               5:
                   "PopUps_DB".Buffer_Cnv_Settings_1 := "Settings_DB".LCnv_Sys[4].Cnv_Level[5].Cnv1;
                   "PopUps_DB".ECnv_Settings := "Settings_DB".ECnv_Sys[4];
                   "PopUps_DB".Buffer_Cnv_Settings_2 := "Settings_DB".LCnv_Sys[4].Cnv_Level[5].Cnv2;
               6:
                   "PopUps_DB".Buffer_Cnv_Settings_1 := "Settings_DB".LCnv_Sys[4].Cnv_Level[6].Cnv1;
                   "PopUps_DB".ECnv_Settings := "Settings_DB".ECnv_Sys[4];
                   "PopUps_DB".Buffer_Cnv_Settings_2 := "Settings_DB".LCnv_Sys[4].Cnv_Level[6].Cnv2;
               7:
                   "PopUps_DB".Buffer_Cnv_Settings_1 := "Settings_DB".LCnv_Sys[4].Cnv_Level[7].Cnv1;
                   "PopUps_DB".ECnv_Settings := "Settings_DB".ECnv_Sys[4];
                   "PopUps_DB".Buffer_Cnv_Settings_2 := "Settings_DB".LCnv_Sys[4].Cnv_Level[7].Cnv2;
               8:
                   "PopUps_DB".Buffer_Cnv_Settings_1 := "Settings_DB".LCnv_Sys[4].Cnv_Level[8].Cnv1;
                   "PopUps_DB".ECnv_Settings := "Settings_DB".ECnv_Sys[4];
                   "PopUps_DB".Buffer_Cnv_Settings_2 := "Settings_DB".LCnv_Sys[4].Cnv_Level[8].Cnv2;
           END_CASE;
       5: //SYSTEM 5
           CASE "CNV_Level_Selected" OF
               1:
                   "PopUps_DB".Buffer_Cnv_Settings_1 := "Settings_DB".LCnv_Sys[5].Cnv_Level[1].Cnv1;
                   "PopUps_DB".ECnv_Settings := "Settings_DB".ECnv_Sys[5];
                   "PopUps_DB".Buffer_Cnv_Settings_2 := "Settings_DB".LCnv_Sys[5].Cnv_Level[1].Cnv2;
               2:
                   "PopUps_DB".Buffer_Cnv_Settings_1 := "Settings_DB".LCnv_Sys[5].Cnv_Level[2].Cnv1;
                   "PopUps_DB".ECnv_Settings := "Settings_DB".ECnv_Sys[5];
                   "PopUps_DB".Buffer_Cnv_Settings_2 := "Settings_DB".LCnv_Sys[5].Cnv_Level[2].Cnv2;
               3:
                   "PopUps_DB".Buffer_Cnv_Settings_1 := "Settings_DB".LCnv_Sys[5].Cnv_Level[3].Cnv1;
                   "PopUps_DB".ECnv_Settings := "Settings_DB".ECnv_Sys[5];
                   "PopUps_DB".Buffer_Cnv_Settings_2 := "Settings_DB".LCnv_Sys[5].Cnv_Level[3].Cnv2;
               4:
                   "PopUps_DB".Buffer_Cnv_Settings_1 := "Settings_DB".LCnv_Sys[5].Cnv_Level[4].Cnv1;
                   "PopUps_DB".ECnv_Settings := "Settings_DB".ECnv_Sys[5];
                   "PopUps_DB".Buffer_Cnv_Settings_2 := "Settings_DB".LCnv_Sys[5].Cnv_Level[4].Cnv2;
               5:
                   "PopUps_DB".Buffer_Cnv_Settings_1 := "Settings_DB".LCnv_Sys[5].Cnv_Level[5].Cnv1;
                   "PopUps_DB".ECnv_Settings := "Settings_DB".ECnv_Sys[5];
                   "PopUps_DB".Buffer_Cnv_Settings_2 := "Settings_DB".LCnv_Sys[5].Cnv_Level[5].Cnv2;
               6:
                   "PopUps_DB".Buffer_Cnv_Settings_1 := "Settings_DB".LCnv_Sys[5].Cnv_Level[6].Cnv1;
                   "PopUps_DB".ECnv_Settings := "Settings_DB".ECnv_Sys[5];
                   "PopUps_DB".Buffer_Cnv_Settings_2 := "Settings_DB".LCnv_Sys[5].Cnv_Level[6].Cnv2;
               7:
                   "PopUps_DB".Buffer_Cnv_Settings_1 := "Settings_DB".LCnv_Sys[5].Cnv_Level[7].Cnv1;
                   "PopUps_DB".ECnv_Settings := "Settings_DB".ECnv_Sys[5];
                   "PopUps_DB".Buffer_Cnv_Settings_2 := "Settings_DB".LCnv_Sys[5].Cnv_Level[7].Cnv2;
               8:
                   "PopUps_DB".Buffer_Cnv_Settings_1 := "Settings_DB".LCnv_Sys[5].Cnv_Level[8].Cnv1;
                   "PopUps_DB".ECnv_Settings := "Settings_DB".ECnv_Sys[5];
                   "PopUps_DB".Buffer_Cnv_Settings_2 := "Settings_DB".LCnv_Sys[5].Cnv_Level[8].Cnv2;
           END_CASE;
   END_CASE;
END_FUNCTION

FUNCTION "CNV_Charge_Settings_FC_1" : Void   // FC59, SCL
{ S7_Optimized_Access := 'TRUE' }
VERSION : 0.1
// stored: AutoNumber true, IsIECCheckEnabled false, SetENOAutomatically false, UDAEnableTagReadback false
   VAR_INPUT
      Sys_No : UInt;
      HMI_Box : UInt;
   END_VAR
   VAR_TEMP
      Level : UInt;
   END_VAR
BEGIN
   #Level := #HMI_Box MOD 10;
   "PopUps_DB_1"."ECnv_Settings"[#Sys_No] := "Settings_DB".ECnv_Sys[#Sys_No];

   CASE #Level OF
       1:
           "PopUps_DB_1"."Buffer_Cnv_Settings_1"[#Sys_No] := "Settings_DB".LCnv_Sys[#Sys_No].Cnv_Level[1].Cnv1;
           "PopUps_DB_1"."Buffer_Cnv_Settings_2"[#Sys_No] := "Settings_DB".LCnv_Sys[#Sys_No].Cnv_Level[1].Cnv2;
       2:
           "PopUps_DB_1"."Buffer_Cnv_Settings_1"[#Sys_No] := "Settings_DB".LCnv_Sys[#Sys_No].Cnv_Level[2].Cnv1;
           "PopUps_DB_1"."Buffer_Cnv_Settings_2"[#Sys_No] := "Settings_DB".LCnv_Sys[#Sys_No].Cnv_Level[2].Cnv2;
       3:
           "PopUps_DB_1"."Buffer_Cnv_Settings_1"[#Sys_No] := "Settings_DB".LCnv_Sys[#Sys_No].Cnv_Level[3].Cnv1;
           "PopUps_DB_1"."Buffer_Cnv_Settings_2"[#Sys_No] := "Settings_DB".LCnv_Sys[#Sys_No].Cnv_Level[3].Cnv2;
       4:
           "PopUps_DB_1"."Buffer_Cnv_Settings_1"[#Sys_No] := "Settings_DB".LCnv_Sys[#Sys_No].Cnv_Level[4].Cnv1;
           "PopUps_DB_1"."Buffer_Cnv_Settings_2"[#Sys_No] := "Settings_DB".LCnv_Sys[#Sys_No].Cnv_Level[4].Cnv2;
       5:
           "PopUps_DB_1"."Buffer_Cnv_Settings_1"[#Sys_No] := "Settings_DB".LCnv_Sys[#Sys_No].Cnv_Level[5].Cnv1;
           "PopUps_DB_1"."Buffer_Cnv_Settings_2"[#Sys_No] := "Settings_DB".LCnv_Sys[#Sys_No].Cnv_Level[5].Cnv2;
       6:
           "PopUps_DB_1"."Buffer_Cnv_Settings_1"[#Sys_No] := "Settings_DB".LCnv_Sys[#Sys_No].Cnv_Level[6].Cnv1;
           "PopUps_DB_1"."Buffer_Cnv_Settings_2"[#Sys_No] := "Settings_DB".LCnv_Sys[#Sys_No].Cnv_Level[6].Cnv2;
       7:
           "PopUps_DB_1"."Buffer_Cnv_Settings_1"[#Sys_No] := "Settings_DB".LCnv_Sys[#Sys_No].Cnv_Level[7].Cnv1;
           "PopUps_DB_1"."Buffer_Cnv_Settings_2"[#Sys_No] := "Settings_DB".LCnv_Sys[#Sys_No].Cnv_Level[7].Cnv2;
       8:
           "PopUps_DB_1"."Buffer_Cnv_Settings_1"[#Sys_No] := "Settings_DB".LCnv_Sys[#Sys_No].Cnv_Level[8].Cnv1;
           "PopUps_DB_1"."Buffer_Cnv_Settings_2"[#Sys_No] := "Settings_DB".LCnv_Sys[#Sys_No].Cnv_Level[8].Cnv2;
   END_CASE;
END_FUNCTION

FUNCTION "CNV_Order_FC" : Void   // FC46, SCL
{ S7_Optimized_Access := 'TRUE' }
VERSION : 0.1
// stored: AutoNumber true, IsIECCheckEnabled false, SetENOAutomatically false, UDAEnableTagReadback false
   VAR_INPUT
      i_Sys : UInt;
      Level : UInt;
      Tower : UInt;
      Transfer_From_To : Byte;
      Pallet_Type : Char;
      Pallet_Allignment : Char;
      Device : String;
      Task_Type : Int;
   END_VAR
   VAR_IN_OUT
      StepTable_0 : "OrderTable_UDT";
   END_VAR
   VAR_TEMP
      StrSys : String;
      StrLev : String;
      Concat1 : String;
      Concat2 : String;
      Source_Location : DInt;
      Destination_Location : DInt;
      Concat3 : String;
      Concat4 : String;
      StrSource : String;
      StrDestination : String;
   END_VAR
BEGIN
   #StrSys := UINT_TO_STRING(#i_Sys);

   // Remove "+"
   IF #StrSys[1] = '+' THEN
       #StrSys := RIGHT(IN := #StrSys, L := LEN(#StrSys) - 1);
   END_IF;

   #StrLev := UINT_TO_STRING(#Level);

   // Remove "+"
   IF #StrLev[1] = '+' THEN
       #StrLev := RIGHT(IN := #StrLev, L := LEN(#StrLev) - 1);
   END_IF;

   IF #Tower = 1 AND #Transfer_From_To = 2 THEN//EXTRACTOR TO CONVEYOR 1
       #StrSource := '120';
       #StrDestination := '100';
   ELSIF #Tower = 2 AND #Transfer_From_To = 2 THEN //EXTRACTOR TO CONVEYOR 2
       #StrSource := '120';
       #StrDestination := '110';
   ELSIF #Tower = 1 AND #Transfer_From_To = 1 THEN //CONVEYOR 1 TO EXTRACTOR
       #StrSource := '100';
       #StrDestination := '120';
   ELSIF #Tower = 2 AND #Transfer_From_To = 1 THEN //CONVEYOR 2 TO EXTRACTOR
       #StrSource := '110';
       #StrDestination := '120';
   ELSIF #Tower = 1 AND #Transfer_From_To = 3 THEN //LOGISTEX TO CONVEYOR 1
       #StrSource := '0';
       #StrDestination := '100';
   ELSIF #Tower = 2 AND #Transfer_From_To = 4 THEN // CONVEYOR 2 TO LOGISTEX
       #StrSource := '110';
       #StrDestination := '0';
   END_IF;

   // Build Source Location
   #Concat1 := CONCAT(IN1 := #StrSource, IN2 := #StrLev);
   #Concat2 := CONCAT(IN1 := #Concat1, IN2 := '0');
   #Source_Location := STRING_TO_DINT(IN := CONCAT(IN1 := #Concat2, IN2 := #StrSys));

   // Build Destinarion Location
   #Concat3 := CONCAT(IN1 := #StrDestination, IN2 := #StrLev);
   #Concat4 := CONCAT(IN1 := #Concat3, IN2 := '0');
   #Destination_Location := STRING_TO_DINT(IN := CONCAT(IN1 := #Concat4, IN2 := #StrSys));

   "Feed_Steptable_FC"(CurrentTime := "Time".CurrentLocalTime,
                       Task_Type := #Task_Type,
                       Source_Location := #Source_Location,
                       Destination_Location := #Destination_Location,
                       Pallet_Type := #Pallet_Type,
                       Pallet_Alignment := #Pallet_Allignment,
                       Shuttle_ID:=0,
                       StepTable := #StepTable_0);
END_FUNCTION

FUNCTION "CNV_Selector" : Void   // FC8, SCL
{ S7_Optimized_Access := 'TRUE' }
VERSION : 0.1
// stored: AutoNumber true, IsIECCheckEnabled false, SetENOAutomatically false, UDAEnableTagReadback false
BEGIN
   //CNV SCREEN SELECTION

   CASE "CNV_System_Selected" OF
       0:
           "CNV_ID_HMI" := 0;
           "CNV_ID_HMI(1)" := 0;

       1://SYSTEM 1
           "CNV_ID_HMI" := "Settings_DB".ECnv_Sys[1].ID; // EXTRACTOR CONVEYOR
           "CNV_HMI".CNV2_Selected[1] := "CNV2_Selected";
           CASE "CNV_Level_Selected" OF
               1: //LEVEL 1
                   IF "CNV2_Selected" = 1 THEN
                       "CNV_ID_HMI(1)" := "Settings_DB".LCnv_Sys[1].Cnv_Level[1].Cnv1.ID; //CNV 1
                   ELSIF "CNV2_Selected" = 2 THEN
                       "CNV_ID_HMI(1)" := "Settings_DB".LCnv_Sys[1].Cnv_Level[1].Cnv2.ID; //CNV 2
                   END_IF;
               2: //LEVEL 2
                   IF "CNV2_Selected" = 1 THEN
                       "CNV_ID_HMI(1)" := "Settings_DB".LCnv_Sys[1].Cnv_Level[2].Cnv1.ID; //CNV 1
                   ELSIF "CNV2_Selected" = 2 THEN
                       "CNV_ID_HMI(1)" := "Settings_DB".LCnv_Sys[1].Cnv_Level[2].Cnv2.ID; //CNV 2
                   END_IF;
               3: //LEVEL 3
                   IF "CNV2_Selected" = 1 THEN
                       "CNV_ID_HMI(1)" := "Settings_DB".LCnv_Sys[1].Cnv_Level[3].Cnv1.ID; //CNV 1
                   ELSIF "CNV2_Selected" = 2 THEN
                       "CNV_ID_HMI(1)" := "Settings_DB".LCnv_Sys[1].Cnv_Level[3].Cnv2.ID; //CNV 2
                   END_IF;
               4: //LEVEL 4
                   IF "CNV2_Selected" = 1 THEN
                       "CNV_ID_HMI(1)" := "Settings_DB".LCnv_Sys[1].Cnv_Level[4].Cnv1.ID; //CNV 1
                   ELSIF "CNV2_Selected" = 2 THEN
                       "CNV_ID_HMI(1)" := "Settings_DB".LCnv_Sys[1].Cnv_Level[4].Cnv2.ID; //CNV 2
                   END_IF;
               5: //LEVEL 5
                   IF "CNV2_Selected" = 1 THEN
                       "CNV_ID_HMI(1)" := "Settings_DB".LCnv_Sys[1].Cnv_Level[5].Cnv1.ID; //CNV 1
                   ELSIF "CNV2_Selected" = 2 THEN
                       "CNV_ID_HMI(1)" := "Settings_DB".LCnv_Sys[1].Cnv_Level[5].Cnv2.ID; //CNV 2
                   END_IF;
               6: //LEVEL 6
                   IF "CNV2_Selected" = 1 THEN
                       "CNV_ID_HMI(1)" := "Settings_DB".LCnv_Sys[1].Cnv_Level[6].Cnv1.ID; //CNV 1
                   ELSIF "CNV2_Selected" = 2 THEN
                       "CNV_ID_HMI(1)" := "Settings_DB".LCnv_Sys[1].Cnv_Level[6].Cnv2.ID; //CNV 2
                   END_IF;
               7: //LEVEL 7
                   IF "CNV2_Selected" = 1 THEN
                       "CNV_ID_HMI(1)" := "Settings_DB".LCnv_Sys[1].Cnv_Level[7].Cnv1.ID; //CNV 1
                   ELSIF "CNV2_Selected" = 2 THEN
                       "CNV_ID_HMI(1)" := "Settings_DB".LCnv_Sys[1].Cnv_Level[7].Cnv2.ID; //CNV 2
                   END_IF;
               8: //LEVEL 8
                   IF "CNV2_Selected" = 1 THEN
                       "CNV_ID_HMI(1)" := "Settings_DB".LCnv_Sys[1].Cnv_Level[8].Cnv1.ID; //CNV 1
                   ELSIF "CNV2_Selected" = 2 THEN
                       "CNV_ID_HMI(1)" := "Settings_DB".LCnv_Sys[1].Cnv_Level[8].Cnv2.ID; //CNV 2
                   END_IF;
           END_CASE;

       2://SYSTEM 2
           "CNV_ID_HMI" := "Settings_DB".ECnv_Sys[2].ID; // EXTRACTOR CONVEYOR
           "CNV_HMI".CNV2_Selected[2] := "CNV2_Selected";
           CASE "CNV_Level_Selected" OF
               1: //LEVEL 1
                   IF "CNV2_Selected" = 1 THEN
                       "CNV_ID_HMI(1)" := "Settings_DB".LCnv_Sys[2].Cnv_Level[1].Cnv1.ID; //CNV 1
                   ELSIF "CNV2_Selected" = 2 THEN
                       "CNV_ID_HMI(1)" := "Settings_DB".LCnv_Sys[2].Cnv_Level[1].Cnv2.ID; //CNV 2
                   END_IF;
               2: //LEVEL 2
                   IF "CNV2_Selected" = 1 THEN
                       "CNV_ID_HMI(1)" := "Settings_DB".LCnv_Sys[2].Cnv_Level[2].Cnv1.ID; //CNV 1
                   ELSIF "CNV2_Selected" = 2 THEN
                       "CNV_ID_HMI(1)" := "Settings_DB".LCnv_Sys[2].Cnv_Level[2].Cnv2.ID; //CNV 2
                   END_IF;
               3: //LEVEL 3
                   IF "CNV2_Selected" = 1 THEN
                       "CNV_ID_HMI(1)" := "Settings_DB".LCnv_Sys[2].Cnv_Level[3].Cnv1.ID; //CNV 1
                   ELSIF "CNV2_Selected" = 2 THEN
                       "CNV_ID_HMI(1)" := "Settings_DB".LCnv_Sys[2].Cnv_Level[3].Cnv2.ID; //CNV 2
                   END_IF;
               4: //LEVEL 4
                   IF "CNV2_Selected" = 1 THEN
                       "CNV_ID_HMI(1)" := "Settings_DB".LCnv_Sys[2].Cnv_Level[4].Cnv1.ID; //CNV 1
                   ELSIF "CNV2_Selected" = 2 THEN
                       "CNV_ID_HMI(1)" := "Settings_DB".LCnv_Sys[2].Cnv_Level[4].Cnv2.ID; //CNV 2
                   END_IF;
               5: //LEVEL 5
                   IF "CNV2_Selected" = 1 THEN
                       "CNV_ID_HMI(1)" := "Settings_DB".LCnv_Sys[2].Cnv_Level[5].Cnv1.ID; //CNV 1
                   ELSIF "CNV2_Selected" = 2 THEN
                       "CNV_ID_HMI(1)" := "Settings_DB".LCnv_Sys[2].Cnv_Level[5].Cnv2.ID; //CNV 2
                   END_IF;
               6: //LEVEL 6
                   IF "CNV2_Selected" = 1 THEN
                       "CNV_ID_HMI(1)" := "Settings_DB".LCnv_Sys[2].Cnv_Level[6].Cnv1.ID; //CNV 1
                   ELSIF "CNV2_Selected" = 2 THEN
                       "CNV_ID_HMI(1)" := "Settings_DB".LCnv_Sys[2].Cnv_Level[6].Cnv2.ID; //CNV 2
                   END_IF;
               7: //LEVEL 7
                   IF "CNV2_Selected" = 1 THEN
                       "CNV_ID_HMI(1)" := "Settings_DB".LCnv_Sys[2].Cnv_Level[7].Cnv1.ID; //CNV 1
                   ELSIF "CNV2_Selected" = 2 THEN
                       "CNV_ID_HMI(1)" := "Settings_DB".LCnv_Sys[2].Cnv_Level[7].Cnv2.ID; //CNV 2
                   END_IF;
               8: //LEVEL 8
                   IF "CNV2_Selected" = 1 THEN
                       "CNV_ID_HMI(1)" := "Settings_DB".LCnv_Sys[2].Cnv_Level[8].Cnv1.ID; //CNV 1
                   ELSIF "CNV2_Selected" = 2 THEN
                       "CNV_ID_HMI(1)" := "Settings_DB".LCnv_Sys[2].Cnv_Level[8].Cnv2.ID; //CNV 2
                   END_IF;
           END_CASE;

       3://SYSTEM 3
           "CNV_ID_HMI" := "Settings_DB".ECnv_Sys[3].ID; // EXTRACTOR CONVEYOR
           "CNV_HMI".CNV2_Selected[3] := "CNV2_Selected";
           CASE "CNV_Level_Selected" OF
               1: //LEVEL 1
                   IF "CNV2_Selected" = 1 THEN
                       "CNV_ID_HMI(1)" := "Settings_DB".LCnv_Sys[3].Cnv_Level[1].Cnv1.ID; //CNV 1
                   ELSIF "CNV2_Selected" = 2 THEN
                       "CNV_ID_HMI(1)" := "Settings_DB".LCnv_Sys[3].Cnv_Level[1].Cnv2.ID; //CNV 2
                   END_IF;
               2: //LEVEL 2
                   IF "CNV2_Selected" = 1 THEN
                       "CNV_ID_HMI(1)" := "Settings_DB".LCnv_Sys[3].Cnv_Level[2].Cnv1.ID; //CNV 1
                   ELSIF "CNV2_Selected" = 2 THEN
                       "CNV_ID_HMI(1)" := "Settings_DB".LCnv_Sys[3].Cnv_Level[2].Cnv2.ID; //CNV 2
                   END_IF;
               3: //LEVEL 3
                   IF "CNV2_Selected" = 1 THEN
                       "CNV_ID_HMI(1)" := "Settings_DB".LCnv_Sys[3].Cnv_Level[3].Cnv1.ID; //CNV 1
                   ELSIF "CNV2_Selected" = 2 THEN
                       "CNV_ID_HMI(1)" := "Settings_DB".LCnv_Sys[3].Cnv_Level[3].Cnv2.ID; //CNV 2
                   END_IF;
               4: //LEVEL 4
                   IF "CNV2_Selected" = 1 THEN
                       "CNV_ID_HMI(1)" := "Settings_DB".LCnv_Sys[3].Cnv_Level[4].Cnv1.ID; //CNV 1
                   ELSIF "CNV2_Selected" = 2 THEN
                       "CNV_ID_HMI(1)" := "Settings_DB".LCnv_Sys[3].Cnv_Level[4].Cnv2.ID; //CNV 2
                   END_IF;
               5: //LEVEL 5
                   IF "CNV2_Selected" = 1 THEN
                       "CNV_ID_HMI(1)" := "Settings_DB".LCnv_Sys[3].Cnv_Level[5].Cnv1.ID; //CNV 1
                   ELSIF "CNV2_Selected" = 2 THEN
                       "CNV_ID_HMI(1)" := "Settings_DB".LCnv_Sys[3].Cnv_Level[5].Cnv2.ID; //CNV 2
                   END_IF;
               6: //LEVEL 6
                   IF "CNV2_Selected" = 1 THEN
                       "CNV_ID_HMI(1)" := "Settings_DB".LCnv_Sys[3].Cnv_Level[6].Cnv1.ID; //CNV 1
                   ELSIF "CNV2_Selected" = 2 THEN
                       "CNV_ID_HMI(1)" := "Settings_DB".LCnv_Sys[3].Cnv_Level[6].Cnv2.ID; //CNV 2
                   END_IF;
               7: //LEVEL 7
                   IF "CNV2_Selected" = 1 THEN
                       "CNV_ID_HMI(1)" := "Settings_DB".LCnv_Sys[3].Cnv_Level[7].Cnv1.ID; //CNV 1
                   ELSIF "CNV2_Selected" = 2 THEN
                       "CNV_ID_HMI(1)" := "Settings_DB".LCnv_Sys[3].Cnv_Level[7].Cnv2.ID; //CNV 2
                   END_IF;
               8: //LEVEL 8
                   IF "CNV2_Selected" = 1 THEN
                       "CNV_ID_HMI(1)" := "Settings_DB".LCnv_Sys[3].Cnv_Level[8].Cnv1.ID; //CNV 1
                   ELSIF "CNV2_Selected" = 2 THEN
                       "CNV_ID_HMI(1)" := "Settings_DB".LCnv_Sys[3].Cnv_Level[8].Cnv2.ID; //CNV 2
                   END_IF;
           END_CASE;

       4://SYSTEM 4
           "CNV_ID_HMI" := "Settings_DB".ECnv_Sys[4].ID; // EXTRACTOR CONVEYOR
           "CNV_HMI".CNV2_Selected[4] := "CNV2_Selected";
           CASE "CNV_Level_Selected" OF
               1: //LEVEL 1
                   IF "CNV2_Selected" = 1 THEN
                       "CNV_ID_HMI(1)" := "Settings_DB".LCnv_Sys[4].Cnv_Level[1].Cnv1.ID; //CNV 1
                   ELSIF "CNV2_Selected" = 2 THEN
                       "CNV_ID_HMI(1)" := "Settings_DB".LCnv_Sys[4].Cnv_Level[1].Cnv2.ID; //CNV 2
                   END_IF;
               2: //LEVEL 2
                   IF "CNV2_Selected" = 1 THEN
                       "CNV_ID_HMI(1)" := "Settings_DB".LCnv_Sys[4].Cnv_Level[2].Cnv1.ID; //CNV 1
                   ELSIF "CNV2_Selected" = 2 THEN
                       "CNV_ID_HMI(1)" := "Settings_DB".LCnv_Sys[4].Cnv_Level[2].Cnv2.ID; //CNV 2
                   END_IF;
               3: //LEVEL 3
                   IF "CNV2_Selected" = 1 THEN
                       "CNV_ID_HMI(1)" := "Settings_DB".LCnv_Sys[4].Cnv_Level[3].Cnv1.ID; //CNV 1
                   ELSIF "CNV2_Selected" = 2 THEN
                       "CNV_ID_HMI(1)" := "Settings_DB".LCnv_Sys[4].Cnv_Level[3].Cnv2.ID; //CNV 2
                   END_IF;
               4: //LEVEL 4
                   IF "CNV2_Selected" = 1 THEN
                       "CNV_ID_HMI(1)" := "Settings_DB".LCnv_Sys[4].Cnv_Level[4].Cnv1.ID; //CNV 1
                   ELSIF "CNV2_Selected" = 2 THEN
                       "CNV_ID_HMI(1)" := "Settings_DB".LCnv_Sys[4].Cnv_Level[4].Cnv2.ID; //CNV 2
                   END_IF;
               5: //LEVEL 5
                   IF "CNV2_Selected" = 1 THEN
                       "CNV_ID_HMI(1)" := "Settings_DB".LCnv_Sys[4].Cnv_Level[5].Cnv1.ID; //CNV 1
                   ELSIF "CNV2_Selected" = 2 THEN
                       "CNV_ID_HMI(1)" := "Settings_DB".LCnv_Sys[4].Cnv_Level[5].Cnv2.ID; //CNV 2
                   END_IF;
               6: //LEVEL 6
                   IF "CNV2_Selected" = 1 THEN
                       "CNV_ID_HMI(1)" := "Settings_DB".LCnv_Sys[4].Cnv_Level[6].Cnv1.ID; //CNV 1
                   ELSIF "CNV2_Selected" = 2 THEN
                       "CNV_ID_HMI(1)" := "Settings_DB".LCnv_Sys[4].Cnv_Level[6].Cnv2.ID; //CNV 2
                   END_IF;
               7: //LEVEL 7
                   IF "CNV2_Selected" = 1 THEN
                       "CNV_ID_HMI(1)" := "Settings_DB".LCnv_Sys[4].Cnv_Level[7].Cnv1.ID; //CNV 1
                   ELSIF "CNV2_Selected" = 2 THEN
                       "CNV_ID_HMI(1)" := "Settings_DB".LCnv_Sys[4].Cnv_Level[7].Cnv2.ID; //CNV 2
                   END_IF;
               8: //LEVEL 8
                   IF "CNV2_Selected" = 1 THEN
                       "CNV_ID_HMI(1)" := "Settings_DB".LCnv_Sys[4].Cnv_Level[8].Cnv1.ID; //CNV 1
                   ELSIF "CNV2_Selected" = 2 THEN
                       "CNV_ID_HMI(1)" := "Settings_DB".LCnv_Sys[4].Cnv_Level[8].Cnv2.ID; //CNV 2
                   END_IF;
           END_CASE;

